// TwinCAT 3 PLC project Tc_SML_MOTION_LAYER
// ProgramVersion: 3.1.4026.18
// libraries:
//   Tc2_Standard, * (Beckhoff Automation GmbH)
//   Tc2_System, * (Beckhoff Automation GmbH)
// project tree:
//   / PlcTask.TcTTO
//   POUs/ MAIN.TcPOU, FB_AxisCtrl.TcPOU, FB_IoLink_In.TcPOU, FB_IoLink_Out.TcPOU, FB_Mapping_In.TcPOU, FB_Mapping_Out.TcPOU, FB_S7RTT_OTG.TcPOU, I_Axis.TcIO, SML_Diagnostics.TcPOU, SML_Home.TcPOU, SML_Power.TcPOU, SML_ProfilePosition.TcPOU, SML_ProfileVelocity.TcPOU, SML_ProfileVelocity_Jog.TcPOU, SML_Reset.TcPOU, SML_Status.TcPOU, SML_Stop.TcPOU, SML_TouchProbe.TcPOU, f_GetProgress.TcPOU, f_GetState.TcPOU
//   DUTs/ E_AXIS_CTRL.TcDUT, E_AXIS_STATE.TcDUT, E_PROGRESS.TcDUT, OpenSML_Axis.TcDUT, SML_DiagCode.TcDUT, ST_AXIS_CTRL.TcDUT, ST_AXIS_INFO.TcDUT, ST_AXIS_STATE.TcDUT, ST_CiA402_Status.TcDUT, ST_DriveIn.TcDUT, ST_DriveOut.TcDUT, ST_MOVE_DATA.TcDUT, U_AXIS_CTRL.TcDUT, U_AXIS_INFO.TcDUT, U_AXIS_STATE.TcDUT, U_MOVE_DATA.TcDUT
//   GVLs/ GVL_SML_CONST.TcGVL

CONFIGURATION Tc_SML_MOTION_LAYER
    RESOURCE PLC ON TwinCAT3
        TASK PlcTask(INTERVAL := T#10ms, PRIORITY := 20);
        PROGRAM MAIN WITH PlcTask : MAIN;
    END_RESOURCE
END_CONFIGURATION

// ---- DUTs/E_AXIS_CTRL.TcDUT
(* ============================================================
   E_AXIS_CTRL - Axis command (eCmd) for FB_AxisCtrl
   SML v6 - Level B (new)

   Level-based command enum: the application writes Ctrl.eCmd;
   FB_AxisCtrl routes the command to the corresponding leaf FB.
   One command at a time => no explicit arbiter (the single value
   of eCmd IS the arbiter).

   Analogous to E_AXIS_CTRL of PLC_MOTION_LAYER, but the commands
   map onto SML's CiA402 FBs instead of the Beckhoff MC_*.
   ============================================================ *)

TYPE E_AXIS_CTRL :
(
    AXIS_NULL          := 0,    // no command: holds the current state
    AXIS_ENABLE        := 1,    // enable drive (Power) and stay idle
    AXIS_DISABLE       := 2,    // disable drive
    AXIS_RESET         := 3,    // fault reset (drive + leaf FBs)
    AXIS_HOME          := 4,    // homing
    AXIS_MOVE_ABS      := 5,    // absolute Profile Position
    AXIS_MOVE_REL      := 6,    // relative Profile Position
    AXIS_MOVE_VELOCITY := 7,    // Profile Velocity (signed velocity)
    AXIS_JOG_POS       := 8,    // jog positive (held)
    AXIS_JOG_NEG       := 9,    // jog negative (held)
    AXIS_MOVE_CSP      := 10,   // CSP (mode 8) + OTG toward Data.lrTargetPosition
    AXIS_STOP          := 11    // Halt (controlled deceleration)
) INT;
END_TYPE

// ---- DUTs/E_AXIS_STATE.TcDUT
(* ============================================================
   E_AXIS_STATE - Axis functional state
   SML v6 - Level B (new)

   Values that are multiples of 100 (= PROGRESS_SPAN) so they can
   compose the COMBINED STATE with E_PROGRESS:
       State.eState = E_AXIS_STATE + E_PROGRESS
   E.g.: AXIS_STATE_MOVING (500) + PROGRESS_BUSY (2) = 502.
   Decompose with f_GetState(502)=500, f_GetProgress(502)=2.

   Here Level B finally USES the f_GetState / f_GetProgress
   functions introduced in Level A.
   ============================================================ *)

TYPE E_AXIS_STATE :
(
    AXIS_STATE_NULL     := 0,     // not initialized
    AXIS_STATE_INIT     := 100,   // init / reset in progress
    AXIS_STATE_DISABLED := 200,   // drive disabled
    AXIS_STATE_IDLE     := 300,   // enabled, stopped, ready
    AXIS_STATE_HOMING   := 400,   // homing
    AXIS_STATE_MOVING   := 500,   // Profile Position / CSP
    AXIS_STATE_VELOCITY := 600,   // Profile Velocity / Jog
    AXIS_STATE_STOPPING := 700,   // Halt
    AXIS_STATE_ERROR    := 900    // error
) INT;
END_TYPE

// ---- DUTs/E_PROGRESS.TcDUT
(* ============================================================
   E_PROGRESS - Unified progress for all SML FBs
   SML v5 - Level A (new)

   Common progress vocabulary, readable by application / HMI /
   diagnostics, replacing the ad-hoc iState:INT semantics used by
   the individual FBs.

   PROJECTION (Level A):
     Each FB keeps its own iState state machine unchanged and, at
     the end of the cycle, exposes eProgress:E_PROGRESS by deriving
     it from iState and from its own flags (xError / xDone / ...).
     No state machine is rewritten.

   COMBINED STATE (Level B groundwork):
     A machine state can be encoded as
       functional_state + E_PROGRESS
     with functional_state a multiple of 100 (see f_GetState /
     f_GetProgress). Not used yet in Level A.
   ============================================================ *)

TYPE E_PROGRESS :
(
    PROGRESS_INVALID := 0,   // not initialized / idle, no request
    PROGRESS_INIT    := 1,   // start request received
    PROGRESS_BUSY    := 2,   // processing
    PROGRESS_PREPARE := 3,   // preparing parameters / preconditions
    PROGRESS_STARTUP := 4,   // running the startup phase
    PROGRESS_CHECK   := 5,   // verifying result / advancing index
    PROGRESS_DONE    := 6,   // completed successfully
    PROGRESS_ERROR   := 7    // error (terminal until reset)
) INT;
END_TYPE

// ---- DUTs/OpenSML_Axis.TcDUT
(* ============================================================
   OpenSML_Axis - Extended CiA402 PDO Data Structure
   SML v4 - Merged from OpenSML + Confa variants

   SOFTWARE STRUCT - no AT %Q*/%I* mapping.
   Use SML_TC3Link to bridge this struct to the TwinCAT I/O tree.
   This keeps the library portable across runtimes and testable
   in simulation without hardware.

   COMPLETE PDO SET (all standard CiA402 objects + Touch Probe):

   OUTPUTS (PLC -> Drive):
     0x6040  ControlWord
     0x6060  Modes_of_operation
     0x607A  Target_Position          [encoder counts]
     0x6081  Profile_Velocity         [drive velocity units - PP mode]
     0x60FF  Target_Velocity          [drive velocity units - PV/CSV mode]
     0x6071  Target_Torque            [0.1 % of rated]
     0x6083  Profile_Acceleration     [drive accel units - PP/PV mode]
     0x6084  Profile_Deceleration     [drive accel units - PP/PV mode]
     0x607C  Home_Offset              [encoder counts - set before homing]
     0x60B8  TouchProbe_ControlWord   [latch trigger control]

   INPUTS (Drive -> PLC):
     0x6041  StatusWord
     0x6061  Modes_of_operation_display
     0x6077  Torque_Actual_Value      [0.1 % of rated]
     0x6064  Position_Actual_Value    [encoder counts]
     0x606C  Velocity_Actual_Value    [drive velocity units]
     0x6078  Current_Actual_Value     [0.1 % of rated]
     0x60F4  Following_Error_Actual_Value [encoder counts]
     0x603F  Error_Code               [drive-specific error number]
     0x60FD  Digital_Inputs           [bitmask of physical digital inputs]
     0x60B9  TouchProbe_StatusWord
     0x60BA  TouchProbe_Rising_Value  [encoder counts - latched on rising edge]
     0x60BB  TouchProbe_Falling_Value [encoder counts - latched on falling edge]

   ControlWord key bits (CiA402 sect. 8.1.3):
     Bit 0  Switch On
     Bit 1  Enable Voltage
     Bit 2  Quick Stop     (1 = run, 0 = activate quick-stop - ACTIVE LOW)
     Bit 3  Enable Operation
     Bit 4  Mode-specific  (New Setpoint in PP / Start Homing in HM)
     Bit 5  Change Setpoint Immediately - blend moves (PP)
     Bit 6  Relative mode  (PP: 0 = absolute, 1 = relative)
     Bit 7  Fault Reset    (rising edge 0->1 clears fault)
     Bit 8  Halt           (1 = decelerate and hold, stay in OperationEnabled)

   StatusWord key bits (CiA402 sect. 8.1.3):
     Bit 0   Ready to Switch On
     Bit 1   Switched On
     Bit 2   Operation Enabled
     Bit 3   Fault
     Bit 4   Voltage Enabled
     Bit 5   Quick Stop     (0 = quick-stop active)
     Bit 6   Switch On Disabled
     Bit 7   Warning
     Bit 9   Remote
     Bit 10  Target Reached / At Velocity / Setpoint Ack (mode-dependent)
     Bit 11  Internal Limit Active
     Bit 12  Mode-specific  (Setpoint Acknowledge in PP / Home Attained in HM)
     Bit 13  Following Error
     Bit 14  Drive-specific (Standstill on many drives)
   ============================================================ *)

TYPE OpenSML_Axis :
STRUCT
    // --- Outputs: PLC -> Drive --------------------------------
    ControlWord          : UINT;   // 0x6040
    Modes_of_operation   : SINT;   // 0x6060
    Target_Position      : DINT;   // 0x607A [encoder counts]
    Profile_Velocity     : UDINT;  // 0x6081 [drive velocity units - PP move speed]
    Target_Velocity      : DINT;   // 0x60FF [drive velocity units - PV/CSV]
    Target_Torque        : INT;    // 0x6071 [0.1 % of rated]
    Profile_Acceleration : UDINT;  // 0x6083 [drive accel units]
    Profile_Deceleration : UDINT;  // 0x6084 [drive accel units]
    Home_Offset          : DINT;   // 0x607C [encoder counts - offset after homing]
    TouchProbe_ControlWord : UINT; // 0x60B8

    // --- Inputs: Drive -> PLC ---------------------------------
    StatusWord                   : UINT;  // 0x6041
    Modes_of_operation_display   : SINT;  // 0x6061
    Torque_Actual_Value          : INT;   // 0x6077 [0.1 % of rated]
    Position_Actual_Value        : DINT;  // 0x6064 [encoder counts]
    Velocity_Actual_Value        : DINT;  // 0x606C [drive velocity units]
    Current_Actual_Value         : INT;   // 0x6078 [0.1 % of rated]
    Following_Error_Actual_Value : DINT;  // 0x60F4 [encoder counts]
    Error_Code                   : UINT;  // 0x603F [drive error number, 0 = no error]
    Digital_Inputs               : UDINT; // 0x60FD [bitmask of physical DI]
    TouchProbe_StatusWord        : UINT;  // 0x60B9
    TouchProbe_Rising_Value      : DINT;  // 0x60BA [encoder counts]
    TouchProbe_Falling_Value     : DINT;  // 0x60BB [encoder counts]
END_STRUCT
END_TYPE

// ---- DUTs/SML_DiagCode.TcDUT
(* ============================================================
   SML_DiagCode - Diagnostic Code Enumeration
   SML v4 - New in v4 (runtime diagnostics)

   Single categorized code used by SML_Diagnostics for both the
   current condition (DiagCode) and the latched first cause
   (FirstFaultCode).  Backed by UINT so it maps cleanly to an HMI
   tag and to alarm tables.

   RANGES:
     0       OK
     1..9    Warnings (motion continues, attention advised)
     10..19  Drive-level faults (CiA402 StatusWord / Error_Code)
     20..29  Library/motion-FB faults (a sub-FB latched an error)
   ============================================================ *)

TYPE SML_DiagCode :
(
    DIAG_OK               := 0,    // No fault, no warning

    // -- Warnings (1..9) ---------------------------------------
    DIAG_WARNING          := 1,    // CiA402 StatusWord bit 7 (generic warning)
    DIAG_INTERNAL_LIMIT   := 2,    // StatusWord bit 11 (internal limit active)

    // -- Drive-level faults (10..19) ---------------------------
    DIAG_DRIVE_FAULT      := 10,   // StatusWord bit 3 (Fault), no specific code
    DIAG_DRIVE_ERRORCODE  := 11,   // StatusWord bit 3 + Error_Code (0x603F) > 0
    DIAG_QUICK_STOP       := 12,   // QuickStopActive (StatusWord bit 5 = 0)
    DIAG_FOLLOWING_ERROR  := 13,   // StatusWord bit 13 (following error)

    // -- Library / motion-FB faults (20..29) -------------------
    DIAG_POWER_ERROR      := 20,   // SML_Power sequence error
    DIAG_HOME_ERROR       := 21,   // SML_Home error (stall/timeout/abort)
    DIAG_MOVE_ERROR       := 22,   // SML_ProfilePosition error (MoveAbs/MoveHome)
    DIAG_VEL_ERROR        := 23,   // SML_ProfileVelocity error
    DIAG_JOG_ERROR        := 24,   // SML_ProfileVelocity_Jog error
    DIAG_TOUCHPROBE_ERROR := 25,   // SML_TouchProbe error
    DIAG_OTG_ERROR        := 26    // FB_S7RTT_OTG constraint error (invalid limits / cycle time)
) UINT;
END_TYPE

// ---- DUTs/ST_AXIS_CTRL.TcDUT
(* ============================================================
   ST_AXIS_CTRL - Command structure (app -> layer)
   SML v6 - Level B (new)

   The "Ctrl" data contract of the Motion Layer pattern. A flat,
   serializable structure (no pointer/interface inside): accessible
   via ADS symbol or copyable onto a bus (MAPPING groundwork).

   The eCmd command is level-based. Motion parameters live in
   ST_MOVE_DATA ("Data").
   ============================================================ *)

TYPE ST_AXIS_CTRL :
STRUCT
    eCmd           : E_AXIS_CTRL;        // requested command
    xEmergencyStop : BOOL := TRUE;       // TRUE = run / FALSE = quick-stop (CiA402 bit 2)
    xSimulation    : BOOL;               // mirror Target_Position -> Position_Actual_Value

    // -- configuration (rarely changed) -----------------------
    Scale          : LREAL := 4096.0;    // [counts/unit] - must be > 0
    CycleTime      : LREAL := 0.001;     // [s] - must match the task (OTG)
    PositionWindow : LREAL := 0.01;      // in-position deadband [units]
    HomeOffset     : DINT  := 0;         // homing offset [encoder counts] -> 0x607C

    // -- TouchProbe (parallel to motion, not an eCmd) ----------
    xTouchProbeEnable  : BOOL;           // arm the TouchProbe hardware
    xTouchProbeRising  : BOOL;           // arm the latch on the rising edge
    xTouchProbeFalling : BOOL;           // arm the latch on the falling edge
END_STRUCT
END_TYPE

// ---- DUTs/ST_AXIS_INFO.TcDUT
(* ============================================================
   ST_AXIS_INFO - Info structure (layer -> app)
   SML v6 - Level B (new)

   The "Info" data contract. Actual values and axis status bits,
   in user units.
   ============================================================ *)

TYPE ST_AXIS_INFO :
STRUCT
    lrActualPosition : LREAL;    // actual position [units]
    lrActualVelocity : LREAL;    // actual velocity [units/s]
    xEnabled         : BOOL;     // drive in OperationEnabled
    xHomed           : BOOL;     // homing done at least once (latch)
    xMoving          : BOOL;     // axis is moving
    xInPosition      : BOOL;     // within PositionWindow (CSP path)

    // -- full CiA402 decoder (from SML_Status) -----------------
    Status           : ST_CiA402_Status;

    // -- TouchProbe results (from SML_TouchProbe) --------------
    xTouchProbeDoneR       : BOOL;
    xTouchProbeDoneF       : BOOL;
    xTouchProbeBusy        : BOOL;
    xTouchProbeError       : BOOL;
    TouchProbeRisingValue  : DINT;   // [encoder counts]
    TouchProbeFallingValue : DINT;   // [encoder counts]
END_STRUCT
END_TYPE

// ---- DUTs/ST_AXIS_STATE.TcDUT
(* ============================================================
   ST_AXIS_STATE - State structure (layer -> app)
   SML v6 - Level B (new)

   The "State" data contract. Command result + progress.
   eState is the COMBINED STATE (E_AXIS_STATE + E_PROGRESS);
   use f_GetState / f_GetProgress to decompose it.
   ============================================================ *)

TYPE ST_AXIS_STATE :
STRUCT
    eState         : INT;            // combined state = E_AXIS_STATE + E_PROGRESS
    eProgress      : E_PROGRESS;     // progress (handy, already decomposed)
    eCmdActive     : E_AXIS_CTRL;    // command being executed
    xDone          : BOOL;           // current command complete
    xError         : BOOL;           // aggregated error

    // -- diagnostics (from SML_Diagnostics) -------------------
    DiagCode       : SML_DiagCode;
    DiagText       : STRING(80);
    FirstFaultCode : SML_DiagCode;
    FirstFaultText : STRING(80);
END_STRUCT
END_TYPE

// ---- DUTs/ST_CiA402_Status.TcDUT
(* ============================================================
   ST_CiA402_Status - Full CiA402 status decoder
   SML v9 - Level B (new)

   Mirrors the outputs of the SML_Status decoder, made available in
   the data contract as a sub-struct of ST_AXIS_INFO (Info.Status).
   Brings into FB_AxisCtrl the granular status bits that used to be
   exposed only by FB_SML.
   ============================================================ *)

TYPE ST_CiA402_Status :
STRUCT
    // -- CiA402 state machine ----------------------------------
    NotReadyToSwitchOn  : BOOL;
    SwitchOnDisabled    : BOOL;
    ReadyToSwitchOn     : BOOL;
    SwitchedOn          : BOOL;
    OperationEnabled    : BOOL;
    QuickStopActive     : BOOL;
    FaultReactionActive : BOOL;
    Fault               : BOOL;

    // -- general status ----------------------------------------
    Warning             : BOOL;   // bit 7
    TargetReached       : BOOL;   // bit 10 (mode-dependent)
    Halted              : BOOL;
    VoltageEnabled      : BOOL;   // bit 4
    InternalLimit       : BOOL;   // bit 11

    // -- active operating mode ---------------------------------
    ProfilePositionMode : BOOL;   // 1
    ProfileVelocityMode : BOOL;   // 3
    VelocityMode        : BOOL;   // 2 (legacy)
    TorqueProfileMode   : BOOL;   // 4
    HomingMode          : BOOL;   // 6
    SyncPositionMode    : BOOL;   // 8 (CSP)
    SyncVelocityMode    : BOOL;   // 9 (CSV)

    // -- motion ------------------------------------------------
    Moving              : BOOL;
    StandStill          : BOOL;
    Homed               : BOOL;

    // -- error / detail ----------------------------------------
    Err                 : BOOL;   // Error_Code != 0
    ErrId               : UINT;   // 0x603F
    ActTorque           : INT;    // 0x6077 [0.1% of rated]
    FollowingError      : DINT;   // 0x60F4 [encoder counts]
END_STRUCT
END_TYPE

// ---- DUTs/ST_DriveIn.TcDUT
(* ============================================================
   ST_DriveIn - INPUT process image (Drive -> PLC)
   SML v9 - I/O bridge (new)

   The "input" half of OpenSML_Axis, SAME order and same types.
   Used for the I/O bridge: declared AT %I* (mapped to the drive's
   TxPDOs) and copied into GVL_AXIS.Axis[n] before the computation.

   Valid for both CoDeSys and TwinCAT (generic IEC 61131-3 ST).
   ============================================================ *)

TYPE ST_DriveIn :
STRUCT
    StatusWord                   : UINT;   // 0x6041
    Modes_of_operation_display   : SINT;   // 0x6061
    Torque_Actual_Value          : INT;    // 0x6077 [0.1 % rated]
    Position_Actual_Value        : DINT;   // 0x6064 [encoder counts]
    Velocity_Actual_Value        : DINT;   // 0x606C [drive velocity units]
    Current_Actual_Value         : INT;    // 0x6078 [0.1 % rated]
    Following_Error_Actual_Value : DINT;   // 0x60F4 [encoder counts]
    Error_Code                   : UINT;   // 0x603F [0 = no error]
    Digital_Inputs               : UDINT;  // 0x60FD [DI bitmask]
    TouchProbe_StatusWord        : UINT;   // 0x60B9
    TouchProbe_Rising_Value      : DINT;   // 0x60BA [encoder counts]
    TouchProbe_Falling_Value     : DINT;   // 0x60BB [encoder counts]
END_STRUCT
END_TYPE

// ---- DUTs/ST_DriveOut.TcDUT
(* ============================================================
   ST_DriveOut - OUTPUT process image (PLC -> Drive)
   SML v9 - I/O bridge (new)

   The "output" half of OpenSML_Axis, SAME order and same types.
   Used for the I/O bridge: declared AT %Q* (mapped to the drive's
   RxPDOs) and copied from GVL_AXIS.Axis[n] after the computation.

   Valid for both CoDeSys and TwinCAT (generic IEC 61131-3 ST).
   On CoDeSys, as an alternative, you can directly link
   GVL_AXIS.Axis[n].<member> in the I/O Mapping tab (no bridge).
   ============================================================ *)

TYPE ST_DriveOut :
STRUCT
    ControlWord            : UINT;   // 0x6040
    Modes_of_operation     : SINT;   // 0x6060
    Target_Position        : DINT;   // 0x607A [encoder counts]
    Profile_Velocity       : UDINT;  // 0x6081 [drive velocity units - PP]
    Target_Velocity        : DINT;   // 0x60FF [drive velocity units - PV/CSV]
    Target_Torque          : INT;    // 0x6071 [0.1 % rated]
    Profile_Acceleration   : UDINT;  // 0x6083 [drive accel units]
    Profile_Deceleration   : UDINT;  // 0x6084 [drive accel units]
    Home_Offset            : DINT;   // 0x607C [encoder counts]
    TouchProbe_ControlWord : UINT;   // 0x60B8
END_STRUCT
END_TYPE

// ---- DUTs/ST_MOVE_DATA.TcDUT
(* ============================================================
   ST_MOVE_DATA - Setpoints and dynamic limits (app -> layer)
   SML v6 - Level B (new)

   The "Data" data contract. All values are in USER UNITS (LREAL).
   FB_AxisCtrl converts to the drive's raw units via Ctrl.Scale
   before passing them to the leaf FBs (PP/PV/Jog); the CSP/OTG
   path works directly in user units.

   Scaling note: velocity/acceleration scale is assumed equal to
   position scale (multiply by Scale). For drives whose velocity
   units 0x6081/0x60FF differ, refine the conversion in the FB.
   ============================================================ *)

TYPE ST_MOVE_DATA :
STRUCT
    lrTargetPosition : LREAL;              // target [units] for MOVE_ABS/REL/CSP
    lrVelocity       : LREAL := 10.0;      // velocity [units/s]; signed for MOVE_VELOCITY
    lrAcceleration   : LREAL := 1000.0;    // [units/s^2]
    lrDeceleration   : LREAL := 1000.0;    // [units/s^2]
    lrJerk           : LREAL := 10000.0;   // [units/s^3] - CSP/OTG only
END_STRUCT
END_TYPE

// ---- DUTs/U_AXIS_CTRL.TcDUT
(* ============================================================
   U_AXIS_CTRL - Bus UNION for the axis command
   SML v8 - Level B / MAPPING (new)

   Overlay of the same memory block as:
     - stData : ST_AXIS_CTRL   (typed view for the logic)
     - aRaw   : byte block      (raw view for fieldbus mapping)

   Fixed size = MAP_SIZE_CTRL (>= SIZEOF(ST_AXIS_CTRL), checked by
   FB_Mapping_In). Lets you link the element to the process image as
   a struct or as a raw block without changing the mapped size.
   ============================================================ *)

TYPE U_AXIS_CTRL :
UNION
    stData : ST_AXIS_CTRL;
    aRaw   : ARRAY[1..GVL_SML_CONST.MAP_SIZE_CTRL] OF BYTE;
END_UNION
END_TYPE

// ---- DUTs/U_AXIS_INFO.TcDUT
(* ============================================================
   U_AXIS_INFO - Bus UNION for the axis info
   SML v8 - Level B / MAPPING (new)

   stData : ST_AXIS_INFO (typed) / aRaw : byte block (fieldbus).
   Fixed size = MAP_SIZE_INFO (>= SIZEOF(ST_AXIS_INFO)).
   ============================================================ *)

TYPE U_AXIS_INFO :
UNION
    stData : ST_AXIS_INFO;
    aRaw   : ARRAY[1..GVL_SML_CONST.MAP_SIZE_INFO] OF BYTE;
END_UNION
END_TYPE

// ---- DUTs/U_AXIS_STATE.TcDUT
(* ============================================================
   U_AXIS_STATE - Bus UNION for the axis state
   SML v8 - Level B / MAPPING (new)

   stData : ST_AXIS_STATE (typed) / aRaw : byte block (fieldbus).
   Fixed size = MAP_SIZE_STATE (>= SIZEOF(ST_AXIS_STATE)).
   ============================================================ *)

TYPE U_AXIS_STATE :
UNION
    stData : ST_AXIS_STATE;
    aRaw   : ARRAY[1..GVL_SML_CONST.MAP_SIZE_STATE] OF BYTE;
END_UNION
END_TYPE

// ---- DUTs/U_MOVE_DATA.TcDUT
(* ============================================================
   U_MOVE_DATA - Bus UNION for the motion setpoints
   SML v8 - Level B / MAPPING (new)

   stData : ST_MOVE_DATA (typed) / aRaw : byte block (fieldbus).
   Fixed size = MAP_SIZE_DATA (>= SIZEOF(ST_MOVE_DATA)).
   ============================================================ *)

TYPE U_MOVE_DATA :
UNION
    stData : ST_MOVE_DATA;
    aRaw   : ARRAY[1..GVL_SML_CONST.MAP_SIZE_DATA] OF BYTE;
END_UNION
END_TYPE

// ---- GVLs/GVL_SML_CONST.TcGVL
(* ============================================================
   GVL_SML_CONST - LIBRARY constants (invariants)
   SML

   Only constants owned by the library (machine-independent).
   The application configuration (number of axes) lives in GVL_App.MAX_AXIS.
   Qualified reference: GVL_SML_CONST.PROGRESS_SPAN, ...
   ============================================================ *)

{attribute 'qualified_only'}
VAR_GLOBAL CONSTANT
    PROGRESS_SPAN : DINT := 100;   // progress band width in the combined state
                                   // (E_AXIS_STATE values are multiples of this)

    // -- MAPPING: fixed size (bytes) of the bus blocks for the UNIONs --
    // Must be >= SIZEOF of the corresponding struct (checked at runtime
    // by FB_Mapping_In/Out via Check). Fixed for a stable process image
    // on the fieldbus.
    MAP_SIZE_CTRL  : UDINT := 64;    // >= SIZEOF(ST_AXIS_CTRL)
    MAP_SIZE_DATA  : UDINT := 64;    // >= SIZEOF(ST_MOVE_DATA)
    MAP_SIZE_STATE : UDINT := 256;   // >= SIZEOF(ST_AXIS_STATE) (holds 2x STRING(80))
    MAP_SIZE_INFO  : UDINT := 128;   // >= SIZEOF(ST_AXIS_INFO) (with Status + TouchProbe)
END_VAR

// ---- POUs/I_Axis.TcIO
INTERFACE I_Axis

METHOD Enable : E_PROGRESS
VAR_INPUT
END_VAR
END_METHOD

METHOD Disable : E_PROGRESS
VAR_INPUT
END_VAR
END_METHOD

METHOD Reset : E_PROGRESS
VAR_INPUT
END_VAR
END_METHOD

METHOD Home : E_PROGRESS
VAR_INPUT
END_VAR
END_METHOD

METHOD MoveAbsolute : E_PROGRESS
VAR_INPUT
    lrPosition : LREAL;   // [units]
    lrVelocity : LREAL;   // [units/s]
END_VAR
END_METHOD

METHOD MoveRelative : E_PROGRESS
VAR_INPUT
    lrDistance : LREAL;   // [units]
    lrVelocity : LREAL;   // [units/s]
END_VAR
END_METHOD

METHOD MoveVelocity : E_PROGRESS
VAR_INPUT
    lrVelocity : LREAL;   // [units/s] signed
END_VAR
END_METHOD

METHOD Jog : E_PROGRESS
VAR_INPUT
    xForward   : BOOL;
    xReverse   : BOOL;
    lrVelocity : LREAL;   // magnitude [units/s]
END_VAR
END_METHOD

METHOD MoveFollow : E_PROGRESS
VAR_INPUT
    lrPosition : LREAL;   // [units] - online re-targetable
    lrVelocity : LREAL;   // [units/s]
END_VAR
END_METHOD

METHOD Stop : E_PROGRESS
VAR_INPUT
END_VAR
END_METHOD

PROPERTY Position : LREAL
GET
END_GET
END_PROPERTY

PROPERTY Enabled : BOOL
GET
END_GET
END_PROPERTY

END_INTERFACE

// ---- POUs/MAIN.TcPOU
PROGRAM MAIN
VAR
END_VAR

END_PROGRAM

// ---- POUs/FB_Mapping_In.TcPOU
(* ============================================================
   FB_Mapping_In - MAPPING bridge FB: bus -> internal (command)
   SML - Level B / MAPPING (library FB)

   Copies the command/setpoint from the bus UNIONs into the internal
   Ctrl/Data structs, for all axes:
     CtrlBus[].stData -> Ctrl[]   ,   DataBus[].stData -> Data[]
   Call at the START of the task, before the axis loop.

   Reusable: arrays passed by VAR_IN_OUT as ARRAY[*] (variable
   length) - no dependency on MAX_AXIS or on any application GVL. The
   application keeps the bus UNION arrays (e.g. GVL_AXIS_MAP.Ctrl/Data)
   and its enable flag, and instantiates this FB.

   GATE: copies only when xEnable = TRUE.
   Runtime size check: if a struct exceeds its bus block (MAP_SIZE_CTRL/DATA),
   the copy is blocked for safety (resize MAP_SIZE_* in GVL_SML_CONST).
   Precondition: all arrays have the same bounds (one entry per axis).
   ============================================================ *)

FUNCTION_BLOCK FB_Mapping_In
VAR_INPUT
    xEnable : BOOL;   // TRUE = perform the copy; FALSE = bypass
END_VAR
VAR_IN_OUT
    CtrlBus : ARRAY[*] OF U_AXIS_CTRL;   // <- bus command  (.stData)
    DataBus : ARRAY[*] OF U_MOVE_DATA;   // <- bus setpoint (.stData)
    Ctrl    : ARRAY[*] OF ST_AXIS_CTRL;  // -> internal command
    Data    : ARRAY[*] OF ST_MOVE_DATA;  // -> internal setpoint
END_VAR
VAR
    i       : DINT;
    bSizeOk : BOOL;
END_VAR

IF NOT xEnable THEN RETURN; END_IF

// -- Bus block size check (safety) ----------------------------
bSizeOk := (SIZEOF(ST_AXIS_CTRL) <= GVL_SML_CONST.MAP_SIZE_CTRL)
       AND (SIZEOF(ST_MOVE_DATA) <= GVL_SML_CONST.MAP_SIZE_DATA);
IF NOT bSizeOk THEN RETURN; END_IF   // blocked: resize MAP_SIZE_*

// -- Copy bus -> internal -------------------------------------
FOR i := LOWER_BOUND(Ctrl, 1) TO UPPER_BOUND(Ctrl, 1) DO
    Ctrl[i] := CtrlBus[i].stData;
    Data[i] := DataBus[i].stData;
END_FOR

END_FUNCTION_BLOCK

// ---- POUs/FB_AxisCtrl.TcPOU
(* ============================================================
   FB_AxisCtrl - Command-driven axis control FB (Level B)
   SML v6 - new

   Brings the Motion Layer pattern of PLC_MOTION_LAYER onto SML:
   instead of wrapping the Beckhoff MC_*, this FB drives DIRECTLY
   SML's CiA402 leaf FBs (Power/Home/ProfilePosition/ProfileVelocity/
   Jog/Stop) + the CSP path with FB_S7RTT_OTG.

   SUPERSET of FB_SML (v9): it also integrates the full status decoder
   SML_Status (-> Info.Status, all CiA402 bits) and SML_TouchProbe
   (-> Info.xTouchProbe* fields, commanded via Ctrl.xTouchProbe* inputs). The TouchProbe
   is PARALLEL to motion (it is not an eCmd) and its error feeds the
   diagnostics but NOT the combined motion state (eState).

   INPUTS / OUTPUTS via the data contract (VAR_IN_OUT):
     Axis  : OpenSML_Axis   drive PDO image
     Ctrl  : ST_AXIS_CTRL   command (eCmd) + config             (app -> layer)
     Data  : ST_MOVE_DATA   motion setpoints [user units]       (app -> layer)
     State : ST_AXIS_STATE  result + combined state            (layer -> app)
     Info  : ST_AXIS_INFO   actual values + bits                (layer -> app)

   ARBITRATION: eCmd is a single value => only one motion command
   active per cycle. No explicit arbiter (unlike FB_SML).

   ENTRY-POINT: call cyclically. As an alternative to writing
   Ctrl.eCmd, you can use the I_Axis methods (equivalent setters).

   IMPLEMENTS I_Axis.
   ============================================================ *)

FUNCTION_BLOCK FB_AxisCtrl IMPLEMENTS I_Axis
VAR_IN_OUT
    Axis  : OpenSML_Axis;
    Ctrl  : ST_AXIS_CTRL;
    Data  : ST_MOVE_DATA;
    State : ST_AXIS_STATE;
    Info  : ST_AXIS_INFO;
END_VAR
VAR
    // -- leaf FBs (execution level, in place of the MC_*) ------
    inst_Power   : SML_Power;
    inst_Reset   : SML_Reset;
    inst_Home    : SML_Home;
    inst_MoveAbs : SML_ProfilePosition;
    inst_MoveVel : SML_ProfileVelocity;
    inst_Jog     : SML_ProfileVelocity_Jog;
    inst_Stop       : SML_Stop;
    inst_Diag       : SML_Diagnostics;
    inst_Status     : SML_Status;         // full CiA402 decoder (superset of FB_SML)
    inst_TouchProbe : SML_TouchProbe;     // TouchProbe (parallel to motion)
    otg          : FB_S7RTT_OTG;

    // -- command -----------------------------------------------
    _eCmd, _eCmdOld : E_AXIS_CTRL;

    // -- latch / pulse ----------------------------------------
    _bEnableReq  : BOOL;       // enable request (ENABLE/DISABLE)
    _xReset      : BOOL;       // reset active (level)
    _xHomedLatch : BOOL;       // homing done at least once
    _eCspState   : INT;        // CSP sub-state: 0 seed, 1 run

    // -- unit conversions (user -> raw drive) -----------------
    _diPos   : DINT;
    _diVelSg : DINT;           // signed velocity (PV)
    _diVelMg : DINT;           // magnitude (Jog)
    _udiVel  : UDINT;
    _udiAcc  : UDINT;
    _udiDec  : UDINT;

    // -- gate -------------------------------------------------
    _xMotionEnable : BOOL;

    // -- flags from the leaf FBs ------------------------------
    _xEnabled, _xPowerErr                          : BOOL;
    _xResetDone, _xResetErr                        : BOOL;
    _xHomeBusy, _xHomeDone, _xHomeErr              : BOOL;
    _xMoveDone, _xMoveBusy, _xMoveMoving, _xMoveErr: BOOL;
    _xAtVel, _xVelMoving, _xVelErr                 : BOOL;
    _xJogMoving, _xJogErr                          : BOOL;
    _xStopped                                      : BOOL;
    _xTpErr                                        : BOOL;   // TouchProbe error (parallel)
    _xInPos, _xCspErr                              : BOOL;
    _xActiveFault, _xAnyErr                        : BOOL;

    // -- combined-state computation ---------------------------
    _eBase : E_AXIS_STATE;
    _eProg : E_PROGRESS;
END_VAR

//------------------------------------------------------------------------------
// /input + guards
//------------------------------------------------------------------------------
_eCmd := Ctrl.eCmd;

IF Ctrl.Scale = 0.0 THEN Ctrl.Scale := 1.0; END_IF   // divide-by-zero guard

IF Ctrl.xSimulation THEN
    Axis.Position_Actual_Value := Axis.Target_Position;  // mirror in simulation
END_IF

// enable latch: any command != NULL/DISABLE implies enable
IF    _eCmd = AXIS_DISABLE THEN _bEnableReq := FALSE;
ELSIF _eCmd <> AXIS_NULL   THEN _bEnableReq := TRUE;
END_IF

_xReset        := (_eCmd = AXIS_RESET);
_xMotionEnable := _xEnabled AND Ctrl.xEmergencyStop;

// user units -> drive raw units (see scaling note in ST_MOVE_DATA)
_diPos   := LREAL_TO_DINT (Data.lrTargetPosition * Ctrl.Scale);
_diVelSg := LREAL_TO_DINT (Data.lrVelocity       * Ctrl.Scale);
_diVelMg := LREAL_TO_DINT (ABS(Data.lrVelocity)  * Ctrl.Scale);
_udiVel  := LREAL_TO_UDINT(ABS(Data.lrVelocity)  * Ctrl.Scale);
_udiAcc  := LREAL_TO_UDINT(Data.lrAcceleration   * Ctrl.Scale);
_udiDec  := LREAL_TO_UDINT(Data.lrDeceleration   * Ctrl.Scale);
//------------------------------------------------------------------------------
// input + guards/
//------------------------------------------------------------------------------

//------------------------------------------------------------------------------
// /leaf FBs - called every cycle, gated via eCmd (like FB_SML)
//------------------------------------------------------------------------------
inst_Power(
    Axis           := Axis,
    xExecute       := _bEnableReq,
    xEmergencyStop := Ctrl.xEmergencyStop,
    xDone          => _xEnabled,
    xError         => _xPowerErr);

inst_Reset(
    Axis     := Axis,
    xExecute := _xReset,
    xDone    => _xResetDone,
    xError   => _xResetErr);

inst_Home(
    Axis         := Axis,
    xEnable      := _xMotionEnable,
    xExecute     := (_eCmd = AXIS_HOME),
    xReset       := _xReset,
    diHomeOffset := Ctrl.HomeOffset,
    xBusy        => _xHomeBusy,
    xDone        => _xHomeDone,
    xError       => _xHomeErr);
IF _xHomeDone THEN _xHomedLatch := TRUE; END_IF

inst_MoveAbs(
    Axis                   := Axis,
    xEnable                := _xMotionEnable,
    xExecute               := (_eCmd = AXIS_MOVE_ABS) OR (_eCmd = AXIS_MOVE_REL),
    xReset                 := _xReset,
    xContinueMove          := FALSE,
    xRelativeMode          := (_eCmd = AXIS_MOVE_REL),
    diTargetPosition       := _diPos,
    udiProfileVelocity     := _udiVel,
    udiProfileAcceleration := _udiAcc,
    udiProfileDeceleration := _udiDec,
    xDone                  => _xMoveDone,
    xBusy                  => _xMoveBusy,
    xMoving                => _xMoveMoving,
    xError                 => _xMoveErr);

inst_MoveVel(
    Axis                   := Axis,
    xEnable                := _xMotionEnable,
    xExecute               := (_eCmd = AXIS_MOVE_VELOCITY),
    xReset                 := _xReset,
    diTargetVelocity       := _diVelSg,
    udiProfileAcceleration := _udiAcc,
    udiProfileDeceleration := _udiDec,
    xMoving                => _xVelMoving,
    xAtVelocity            => _xAtVel,
    xError                 => _xVelErr);

inst_Jog(
    Axis                   := Axis,
    xEnable                := _xMotionEnable,
    xExecute_Jog_F         := (_eCmd = AXIS_JOG_POS),
    xExecute_Jog_R         := (_eCmd = AXIS_JOG_NEG),
    xReset                 := _xReset,
    diProfileVelocity      := _diVelMg,
    udiProfileAcceleration := _udiAcc,
    udiProfileDeceleration := _udiDec,
    xMoving                => _xJogMoving,
    xError                 => _xJogErr);

inst_Stop(
    Axis     := Axis,
    xStop    := (_eCmd = AXIS_STOP),
    xStopped => _xStopped);

// full CiA402 decoder (read-only) -> Info.Status
inst_Status(
    Axis                       := Axis,
    xEnable                    := TRUE,
    Status_NotReadyToSwitchOn  => Info.Status.NotReadyToSwitchOn,
    Status_SwitchOnDisabled    => Info.Status.SwitchOnDisabled,
    Status_ReadyToSwitchOn     => Info.Status.ReadyToSwitchOn,
    Status_SwitchedOn          => Info.Status.SwitchedOn,
    Status_OperationEnabled    => Info.Status.OperationEnabled,
    Status_QuickStopActive     => Info.Status.QuickStopActive,
    Status_FaultReactionActive => Info.Status.FaultReactionActive,
    Status_Fault               => Info.Status.Fault,
    Status_Warning             => Info.Status.Warning,
    Status_TargetReached       => Info.Status.TargetReached,
    Status_Halted              => Info.Status.Halted,
    Status_VoltageEnabled      => Info.Status.VoltageEnabled,
    Status_InternalLimit       => Info.Status.InternalLimit,
    Status_ProfilePositionMode => Info.Status.ProfilePositionMode,
    Status_ProfileVelocityMode => Info.Status.ProfileVelocityMode,
    Status_VelocityMode        => Info.Status.VelocityMode,
    Status_TorqueProfileMode   => Info.Status.TorqueProfileMode,
    Status_HomingMode          => Info.Status.HomingMode,
    Status_SyncPositionMode    => Info.Status.SyncPositionMode,
    Status_SyncVelocityMode    => Info.Status.SyncVelocityMode,
    Status_Moving              => Info.Status.Moving,
    Status_StandStill          => Info.Status.StandStill,
    Status_Homed               => Info.Status.Homed,
    StatusErr                  => Info.Status.Err,
    ErrId                      => Info.Status.ErrId,
    ActPosition                => ,
    ActSpeed                   => ,
    ActTorque                  => Info.Status.ActTorque,
    FollowingError             => Info.Status.FollowingError);

// TouchProbe (parallel to motion) -> Info.xTouchProbe*
inst_TouchProbe(
    Axis                     := Axis,
    xEnable                  := _xMotionEnable,
    xExecute                 := Ctrl.xTouchProbeEnable,
    xRisingCapture           := Ctrl.xTouchProbeEnable AND Ctrl.xTouchProbeRising,
    xFallingCapture          := Ctrl.xTouchProbeEnable AND Ctrl.xTouchProbeFalling,
    xReset                   := _xReset,
    xDone_R                  => Info.xTouchProbeDoneR,
    xDone_F                  => Info.xTouchProbeDoneF,
    xBusy                    => Info.xTouchProbeBusy,
    xError                   => _xTpErr,
    TouchProbe_Rising_Value  => Info.TouchProbeRisingValue,
    TouchProbe_Falling_Value => Info.TouchProbeFallingValue);
Info.xTouchProbeError := _xTpErr;
//------------------------------------------------------------------------------
// leaf FBs/
//------------------------------------------------------------------------------

//------------------------------------------------------------------------------
// /CSP + OTG - active only with eCmd = AXIS_MOVE_CSP
//------------------------------------------------------------------------------
_xInPos := FALSE;
IF (_eCmd = AXIS_MOVE_CSP) AND _xMotionEnable THEN
    Info.lrActualPosition := DINT_TO_LREAL(Axis.Position_Actual_Value) / Ctrl.Scale;
    CASE _eCspState OF
        0: // switch to CSP (mode 8) + seed OTG at the actual position
            Axis.Modes_of_operation := 8;
            Axis.ControlWord.3      := (Axis.Modes_of_operation_display = 8);
            otg(
                xInit            := TRUE,
                CurrentPosition  := Info.lrActualPosition,
                ControlInterface := TRUE,
                TargetPosition   := Data.lrTargetPosition,
                TargetVelocity   := 0.0,
                CycleTIme        := Ctrl.CycleTime,
                MaxVelocity      := Data.lrVelocity,
                MaxAcceleration  := Data.lrAcceleration,
                MaxJerk          := Data.lrJerk);
            IF (Axis.StatusWord.2 AND Axis.Modes_of_operation_display = 8) OR Ctrl.xSimulation THEN
                _eCspState := 1;
            END_IF

        1: // CSP motion loop
            otg(
                xInit            := FALSE,
                ControlInterface := FALSE,
                TargetPosition   := Data.lrTargetPosition,
                TargetVelocity   := 0.0,
                CycleTIme        := Ctrl.CycleTime,
                MaxVelocity      := Data.lrVelocity,
                MaxAcceleration  := Data.lrAcceleration,
                MaxJerk          := Data.lrJerk);
            Axis.Target_Position := LREAL_TO_DINT(otg.NewPosition * Ctrl.Scale);
            _xInPos := ABS(otg.NewPosition - Data.lrTargetPosition) < Ctrl.PositionWindow;
    END_CASE
    _xCspErr := Axis.StatusWord.13 OR Axis.StatusWord.3 OR otg.xError OR _xPowerErr;
ELSE
    _eCspState := 0;      // reset the sub-state when not in CSP
    _xCspErr   := FALSE;
END_IF
//------------------------------------------------------------------------------
// CSP + OTG/
//------------------------------------------------------------------------------

//------------------------------------------------------------------------------
// /aggregated diagnostics
//------------------------------------------------------------------------------
inst_Diag(
    Axis             := Axis,
    xReset           := _xReset,
    xResetCount      := FALSE,
    xPowerError      := _xPowerErr,
    xHomeError       := _xHomeErr,
    xMoveError       := _xMoveErr,
    xVelError        := _xVelErr,
    xJogError        := _xJogErr,
    xTouchProbeError := _xTpErr,
    xOtgError        := otg.xError,
    DiagCode         => State.DiagCode,
    DiagText         => State.DiagText,
    xActiveFault     => _xActiveFault,
    xActiveWarning   => ,
    FirstFaultCode   => State.FirstFaultCode,
    FirstFaultText   => State.FirstFaultText,
    DriveErrorCode   => ,
    FollowingError   => ,
    FaultCount       => );
//------------------------------------------------------------------------------
// aggregated diagnostics/
//------------------------------------------------------------------------------

//------------------------------------------------------------------------------
// /Info (feedback) + aggregated error
//------------------------------------------------------------------------------
Info.lrActualPosition := DINT_TO_LREAL(Axis.Position_Actual_Value) / Ctrl.Scale;
Info.lrActualVelocity := DINT_TO_LREAL(Axis.Velocity_Actual_Value) / Ctrl.Scale;
Info.xEnabled         := _xEnabled;
Info.xHomed           := _xHomedLatch;
Info.xMoving          := _xMoveMoving OR _xVelMoving OR _xJogMoving OR (_eCmd = AXIS_MOVE_CSP);
Info.xInPosition      := _xInPos;

_xAnyErr := _xPowerErr OR _xHomeErr OR _xMoveErr OR _xVelErr
            OR _xJogErr OR _xCspErr OR _xResetErr;
//------------------------------------------------------------------------------
// Info + error/
//------------------------------------------------------------------------------

//------------------------------------------------------------------------------
// /combined state  eState = E_AXIS_STATE + E_PROGRESS
//------------------------------------------------------------------------------
IF _xAnyErr THEN
    _eBase := AXIS_STATE_ERROR;
    _eProg := PROGRESS_ERROR;
ELSE
    CASE _eCmd OF
        AXIS_NULL:
            IF _xEnabled THEN _eBase := AXIS_STATE_IDLE; ELSE _eBase := AXIS_STATE_DISABLED; END_IF
            _eProg := PROGRESS_INVALID;

        AXIS_ENABLE:
            _eBase := AXIS_STATE_IDLE;
            IF _xEnabled THEN _eProg := PROGRESS_DONE; ELSE _eProg := PROGRESS_BUSY; END_IF

        AXIS_DISABLE:
            _eBase := AXIS_STATE_DISABLED;
            IF _xEnabled THEN _eProg := PROGRESS_BUSY; ELSE _eProg := PROGRESS_DONE; END_IF

        AXIS_RESET:
            _eBase := AXIS_STATE_INIT;
            IF _xResetDone THEN _eProg := PROGRESS_DONE; ELSE _eProg := PROGRESS_BUSY; END_IF

        AXIS_HOME:
            _eBase := AXIS_STATE_HOMING;
            IF _xHomeDone THEN _eProg := PROGRESS_DONE; ELSE _eProg := PROGRESS_BUSY; END_IF

        AXIS_MOVE_ABS, AXIS_MOVE_REL:
            _eBase := AXIS_STATE_MOVING;
            IF _xMoveDone THEN _eProg := PROGRESS_DONE; ELSE _eProg := PROGRESS_BUSY; END_IF

        AXIS_MOVE_CSP:
            _eBase := AXIS_STATE_MOVING;
            IF _xInPos THEN _eProg := PROGRESS_DONE; ELSE _eProg := PROGRESS_BUSY; END_IF

        AXIS_MOVE_VELOCITY:
            _eBase := AXIS_STATE_VELOCITY;
            IF _xAtVel THEN _eProg := PROGRESS_DONE; ELSE _eProg := PROGRESS_BUSY; END_IF

        AXIS_JOG_POS, AXIS_JOG_NEG:
            _eBase := AXIS_STATE_VELOCITY;
            _eProg := PROGRESS_BUSY;      // continuous jog: no discrete DONE

        AXIS_STOP:
            _eBase := AXIS_STATE_STOPPING;
            IF _xStopped THEN _eProg := PROGRESS_DONE; ELSE _eProg := PROGRESS_BUSY; END_IF
    END_CASE
END_IF

State.eProgress  := _eProg;
State.eState     := TO_INT(_eBase) + TO_INT(_eProg);   // combined state
State.eCmdActive := _eCmd;
State.xError     := _xAnyErr;
State.xDone      := (_eProg = PROGRESS_DONE);

_eCmdOld := _eCmd;
//------------------------------------------------------------------------------
// combined state/
//------------------------------------------------------------------------------


(* ============================================================
   METHODS / PROPERTIES of I_Axis
   Real code in  FB_AxisCtrl_METHODS.txt  (to be created as
   METHOD/PROPERTY objects under this FB in CoDeSys).
   They are setters: they set Ctrl.eCmd (+ Data) and return
   State.eProgress.
   ============================================================ *)

METHOD Enable : E_PROGRESS
VAR_INPUT
END_VAR
Ctrl.eCmd := AXIS_ENABLE;
Enable    := State.eProgress;
END_METHOD

METHOD Disable : E_PROGRESS
VAR_INPUT
END_VAR
Ctrl.eCmd := AXIS_DISABLE;
Disable   := State.eProgress;
END_METHOD

METHOD Reset : E_PROGRESS
VAR_INPUT
END_VAR
Ctrl.eCmd := AXIS_RESET;
Reset     := State.eProgress;
END_METHOD

METHOD Home : E_PROGRESS
VAR_INPUT
END_VAR
Ctrl.eCmd := AXIS_HOME;
Home      := State.eProgress;
END_METHOD

METHOD MoveAbsolute : E_PROGRESS
VAR_INPUT
    lrPosition : LREAL;
    lrVelocity : LREAL;
END_VAR
Ctrl.eCmd             := AXIS_MOVE_ABS;
Data.lrTargetPosition := lrPosition;
Data.lrVelocity       := lrVelocity;
MoveAbsolute          := State.eProgress;
END_METHOD

METHOD MoveRelative : E_PROGRESS
VAR_INPUT
    lrDistance : LREAL;
    lrVelocity : LREAL;
END_VAR
Ctrl.eCmd             := AXIS_MOVE_REL;
Data.lrTargetPosition := lrDistance;
Data.lrVelocity       := lrVelocity;
MoveRelative          := State.eProgress;
END_METHOD

METHOD MoveVelocity : E_PROGRESS
VAR_INPUT
    lrVelocity : LREAL;   // signed
END_VAR
Ctrl.eCmd       := AXIS_MOVE_VELOCITY;
Data.lrVelocity := lrVelocity;
MoveVelocity    := State.eProgress;
END_METHOD

METHOD Jog : E_PROGRESS
VAR_INPUT
    xForward   : BOOL;
    xReverse   : BOOL;
    lrVelocity : LREAL;   // magnitudo
END_VAR
IF    xForward THEN Ctrl.eCmd := AXIS_JOG_POS;
ELSIF xReverse THEN Ctrl.eCmd := AXIS_JOG_NEG;
ELSE               Ctrl.eCmd := AXIS_NULL;
END_IF
Data.lrVelocity := lrVelocity;
Jog             := State.eProgress;
END_METHOD

METHOD MoveFollow : E_PROGRESS
VAR_INPUT
    lrPosition : LREAL;
    lrVelocity : LREAL;
END_VAR
Ctrl.eCmd             := AXIS_MOVE_CSP;
Data.lrTargetPosition := lrPosition;
Data.lrVelocity       := lrVelocity;
MoveFollow            := State.eProgress;
END_METHOD

METHOD Stop : E_PROGRESS
VAR_INPUT
END_VAR
Ctrl.eCmd := AXIS_STOP;
Stop      := State.eProgress;
END_METHOD

PROPERTY Position : LREAL
GET
Position := Info.lrActualPosition;
END_GET
END_PROPERTY

PROPERTY Enabled : BOOL
GET
Enabled := Info.xEnabled;
END_GET
END_PROPERTY

END_FUNCTION_BLOCK

// ---- POUs/SML_Power.TcPOU
(* ============================================================
   SML_Power - CiA402 Drive Power-On / Power-Off Sequencer
   SML v4 - Merged (best of OpenSML_Power + SML_Power/Confa)

   Drives the CiA402 state machine:
     SwitchOnDisabled -> ReadyToSwitchOn -> SwitchedOn -> OperationEnabled

   KEY DESIGN CHOICES (vs original OpenSML):
   - xExecute (edge/level) instead of xEnable:
     After a fault reset the drive returns to Idle and REQUIRES a
     new xExecute pulse.  This prevents automatic re-enable after
     any fault - the operator must consciously re-request power.
   - Single tonTimeout instance with explicit IN management per state.
   - Proper CiA402 Shutdown command on disable (bit3=0, bit0=0).
   - All control bits forced low in error state.

   EMERGENCY STOP:
     xEmergencyStop = TRUE  -> ControlWord bit 2 = 1 -> normal run
     xEmergencyStop = FALSE -> ControlWord bit 2 = 0 -> quick-stop
   Applied every cycle regardless of state.
   ============================================================ *)

FUNCTION_BLOCK SML_Power
VAR_IN_OUT
    Axis : OpenSML_Axis;
END_VAR
VAR_INPUT
    xExecute       : BOOL;           // Level/edge: request drive enable; drop to disable
    xEmergencyStop : BOOL := TRUE;   // TRUE = normal run, FALSE = quick-stop (CiA402 bit 2)
END_VAR
VAR_OUTPUT
    xDone  : BOOL; // Drive in OperationEnabled state, ready for motion FBs
    xError : BOOL; // Fault present or power-up sequence timed out
    eProgress : E_PROGRESS; // Level A: unified progress (projection of iState)
END_VAR
VAR
    iState     : INT;
    tonTimeout : TON;
    tTimeOut   : TIME := T#500MS; // Max time allowed per CiA402 state transition
END_VAR

// -- Quick-Stop line - written every scan regardless of state --------------
// CiA402 bit 2: 1 = normal, 0 = quick-stop. Active-LOW - never invert here.
Axis.ControlWord.2 := xEmergencyStop;

// -- Single timer instance - IN assigned per state -------------------------
tonTimeout(PT := tTimeOut);

CASE iState OF

    0: // Idle - safe default; wait for execute request
        xDone  := FALSE;
        xError := FALSE;
        tonTimeout.IN := FALSE;
        Axis.ControlWord.0 := FALSE; // Switch On
        Axis.ControlWord.1 := FALSE; // Enable Voltage
        Axis.ControlWord.3 := FALSE; // Enable Operation
        Axis.ControlWord.7 := FALSE; // Fault Reset (pre-clear)
        IF xExecute THEN
            IF Axis.StatusWord.3 THEN
                iState := 10; // Fault active -> reset first
            ELSE
                iState := 20; // No fault -> begin enable sequence
            END_IF
        END_IF

    10: // Fault Reset - pulse bit 7 (rising edge 0->1 clears fault)
        // On success: return to IDLE (not directly to enable).
        // Operator must re-assert xExecute to intentionally re-enable.
        Axis.ControlWord.7 := TRUE;
        tonTimeout.IN := TRUE;
        IF tonTimeout.Q AND NOT Axis.StatusWord.3 THEN
            Axis.ControlWord.7 := FALSE;
            tonTimeout.IN := FALSE;
            iState := 0; // Back to idle - requires deliberate re-enable
        ELSIF tonTimeout.Q THEN
            tonTimeout.IN := FALSE;
            iState := 999; // Drive did not clear fault within timeout
        END_IF

    20: // Enable Voltage - Shutdown command: bit1=1, bit0=0, bit3=0
        // Transitions: SwitchOnDisabled -> ReadyToSwitchOn
        Axis.ControlWord.1 := TRUE;
        tonTimeout.IN := TRUE;
        IF Axis.StatusWord.0 THEN
            // StatusWord bit 0 = Ready to Switch On confirmed
            tonTimeout.IN := FALSE;
            iState := 30;
        ELSIF tonTimeout.Q THEN
            tonTimeout.IN := FALSE;
            iState := 999;
        END_IF

    30: // Switch On - command: bit1=1, bit0=1, bit3=0
        // Transitions: ReadyToSwitchOn -> SwitchedOn
        Axis.ControlWord.0 := TRUE;
        tonTimeout.IN := TRUE;
        IF Axis.StatusWord.0 AND Axis.StatusWord.1 THEN
            // StatusWord bits 0+1 = Switched On confirmed
            tonTimeout.IN := FALSE;
            iState := 40;
        ELSIF tonTimeout.Q THEN
            tonTimeout.IN := FALSE;
            iState := 999;
        END_IF

    40: // Enable Operation - command: bit0=1, bit1=1, bit3=1
        // Transitions: SwitchedOn -> OperationEnabled
        // Freeze target position BEFORE asserting bit3 to prevent a position jump
        Axis.Target_Position := Axis.Position_Actual_Value;
        Axis.ControlWord.3 := TRUE;
        tonTimeout.IN := TRUE;
        IF Axis.StatusWord.0 AND Axis.StatusWord.1 AND Axis.StatusWord.2 THEN
            // OperationEnabled confirmed
            tonTimeout.IN := FALSE;
            iState := 50;
        ELSIF tonTimeout.Q THEN
            tonTimeout.IN := FALSE;
            iState := 999;
        END_IF

    50: // Running - drive in OperationEnabled, accepting setpoints
        xDone := TRUE;
        IF NOT xExecute THEN
            // CiA402 Shutdown: bit3=0 (Disable Operation) + bit0=0 (Switch Off)
            Axis.ControlWord.3 := FALSE;
            Axis.ControlWord.0 := FALSE;
            iState := 0;
        ELSIF Axis.StatusWord.3 THEN
            // Drive fault while running
            iState := 999;
        ELSIF NOT Axis.StatusWord.5 AND xEmergencyStop THEN
            // M3: QuickStopActive (StatusWord bit 5 = 0) but E-stop has been
            // released (xEmergencyStop = TRUE). Depending on quick-stop option
            // code 0x605A the drive may stay in QuickStopActive and NOT auto-
            // recover. Re-run the enable sequence from Switch-On to bring the
            // drive back to OperationEnabled. xDone drops until re-confirmed.
            xDone := FALSE;
            iState := 20;
        END_IF

    999: // Error - latched; reset by dropping xExecute
        tonTimeout.IN := FALSE;
        xDone  := FALSE;
        xError := TRUE;
        Axis.ControlWord.0 := FALSE; // Force low for safety
        Axis.ControlWord.3 := FALSE;
        IF NOT xExecute THEN
            iState := 0;
        END_IF

END_CASE

// -- Level A: unified progress projection (E_PROGRESS) --------------
IF    xError     THEN eProgress := PROGRESS_ERROR;
ELSIF xDone      THEN eProgress := PROGRESS_DONE;      // OperationEnabled (iState 50)
ELSIF iState = 0 THEN eProgress := PROGRESS_INVALID;   // idle
ELSE                  eProgress := PROGRESS_BUSY;       // sequence in progress
END_IF

END_FUNCTION_BLOCK

// ---- POUs/SML_Reset.TcPOU
(* ============================================================
   SML_Reset - CiA402 Fault Reset (standalone FB)
   SML v4 - Merged (from Confa; not present in original OpenSML)

   Pulses ControlWord bit 7 (rising edge 0->1) to clear a drive
   fault independently of the power sequence.

   Use this FB when you need to reset a fault without going through
   the full SML_Power enable sequence, for example to clear a
   non-critical warning while the drive is in a known safe state.

   State machine:
     0 Idle -> 10 Reset pulse -> 20 Done (wait xExecute drop) -> 0
                             -> 999 Error (fault not cleared)
   ============================================================ *)

FUNCTION_BLOCK SML_Reset
VAR_IN_OUT
    Axis : OpenSML_Axis;
END_VAR
VAR_INPUT
    xExecute : BOOL; // Pulse or level: trigger fault reset
END_VAR
VAR_OUTPUT
    xDone  : BOOL; // Fault cleared successfully
    xError : BOOL; // Fault not cleared within timeout
    eProgress : E_PROGRESS; // Level A: unified progress (projection of iState)
END_VAR
VAR
    iState     : INT;
    tonTimeout : TON;
    tTimeOut   : TIME := T#500MS;
END_VAR

CASE iState OF

    0: // Idle - pre-clear bit 7, wait for execute
        Axis.ControlWord.7 := FALSE; // Rising edge requires bit7 to start at 0
        xDone  := FALSE;
        xError := FALSE;
        IF xExecute THEN
            iState := 10;
        END_IF

    10: // Assert Fault Reset bit (rising edge 0->1)
        Axis.ControlWord.7 := TRUE;
        tonTimeout(IN := TRUE, PT := tTimeOut);
        IF tonTimeout.Q AND NOT Axis.StatusWord.3 THEN
            // Fault cleared
            Axis.ControlWord.7 := FALSE;
            xDone := TRUE;
            tonTimeout(IN := FALSE);
            iState := 20;
        ELSIF tonTimeout.Q THEN
            // Persistent fault - hardware intervention required
            Axis.ControlWord.7 := FALSE;
            tonTimeout(IN := FALSE);
            iState := 999;
        END_IF

    20: // Done - hold until xExecute drops (prevents continuous re-reset)
        IF NOT xExecute THEN
            iState := 0;
        END_IF

    999: // Error - fault not cleared; reset by dropping xExecute
        tonTimeout(IN := FALSE);
        Axis.ControlWord.7 := FALSE;
        xError := TRUE;
        IF NOT xExecute THEN
            iState := 0;
        END_IF

END_CASE

// -- Level A: unified progress projection (E_PROGRESS) --------------
IF    xError     THEN eProgress := PROGRESS_ERROR;
ELSIF xDone      THEN eProgress := PROGRESS_DONE;
ELSIF iState = 0 THEN eProgress := PROGRESS_INVALID;
ELSE                  eProgress := PROGRESS_BUSY;
END_IF

END_FUNCTION_BLOCK

// ---- POUs/SML_Home.TcPOU
(* ============================================================
   SML_Home - CiA402 Homing Sequence (mode 6)
   SML v4 - Merged (OpenSML_Home + SML_Home/Confa)

   Prerequisites - configure via SDO or EtherCAT startup params:
     0x6098  Homing Method
     0x6099.01  Speed for limit switch search
     0x6099.02  Speed for index pulse
     0x609A  Homing Acceleration

   The homing offset (0x607C) is written via PDO at runtime
   through diHomeOffset - no SDO access needed.

   CiA402 completion: StatusWord bit 10 (Target Reached) AND
   bit 12 (Home Attained) must both be set.

   State flow:
     0 Idle -> 10 Mode Switch -> 20 Homing -> 30 Done -> 40 Handshake -> 0
                                         -> 999 Error

   Stall watchdog (state 20): if position doesn't change for
   tStallTimeout, the homing sequence is aborted.
   ============================================================ *)

FUNCTION_BLOCK SML_Home
VAR_IN_OUT
    Axis : OpenSML_Axis;
END_VAR
VAR_INPUT
    xEnable        : BOOL;           // Level: FB active; drop to abort
    xExecute       : BOOL;           // Edge/level: start homing
    xReset         : BOOL;           // Pulse: acknowledge error and return to idle
    diHomeOffset   : DINT;           // Home offset [encoder counts] - written to 0x607C
    tStallTimeout  : TIME := T#10S;  // Max time without position change before error
END_VAR
VAR_OUTPUT
    xBusy  : BOOL; // Homing sequence in progress
    xDone  : BOOL; // Homing completed successfully
    xError : BOOL; // Error: fault, stall, timeout, or operator abort
    eProgress : E_PROGRESS; // Level A: unified progress (projection of iState)
END_VAR
VAR
    iState     : INT;
    tonStall   : TON;  // Stall watchdog
    tonMode    : TON;  // Mode-switch timeout guard
    Pos_Old    : DINT; // Previous-cycle position for stall detection
END_VAR

CASE iState OF

    0: // Idle - reset outputs, capture baseline position for stall detection
        xBusy  := FALSE;
        xDone  := FALSE;
        xError := FALSE;
        tonStall.IN := FALSE;
        tonMode.IN  := FALSE;
        Pos_Old := Axis.Position_Actual_Value; // Baseline so state 20 starts correctly

        IF xEnable THEN
            IF xExecute AND Axis.StatusWord.1         // SwitchedOn
                        AND Axis.StatusWord.2         // OperationEnabled
                        AND Axis.Modes_of_operation_display = 6 // Already in Homing mode
                        AND NOT Axis.StatusWord.3 THEN
                iState := 10;

            ELSIF xExecute AND Axis.StatusWord.1
                           AND Axis.Modes_of_operation_display <> 6 THEN
                // Different mode active - drop EnableOperation for mode switch
                Axis.ControlWord.3 := FALSE;
                iState := 10;

            ELSIF xExecute OR Axis.StatusWord.3 THEN
                iState := 999; // Drive not ready or fault present
            END_IF
        END_IF

    10: // Mode Switch - request Homing mode, write offset, re-enable operation
        tonMode(IN := TRUE, PT := T#2S); // Mode switch should be nearly instantaneous
        Axis.ControlWord.4      := FALSE;       // Clear Start Homing bit before arming
        Axis.Modes_of_operation := 6;           // Request Homing mode
        Axis.Home_Offset        := diHomeOffset; // Write offset to 0x607C via PDO

        // Re-enable operation only when drive confirms mode 6 is active
        Axis.ControlWord.3 := (Axis.Modes_of_operation_display = 6);

        IF Axis.StatusWord.3 OR NOT xEnable OR tonMode.Q THEN
            tonMode.IN := FALSE;
            iState := 999;
        ELSIF Axis.StatusWord.2 AND Axis.ControlWord.3 THEN
            // OperationEnabled confirmed in Homing mode
            tonMode.IN := FALSE;
            xBusy := TRUE;
            iState := 20;
        END_IF

    20: // Homing in progress - arm Start Homing, monitor completion and stall
        Axis.ControlWord.4 := TRUE; // Start Homing (bit 4 in HM mode)

        // Stall watchdog: timer runs while position is unchanged from last cycle.
        // Pos_Old updated AFTER timer call so comparison is current-vs-previous.
        tonStall(IN := (Axis.Position_Actual_Value = Pos_Old), PT := tStallTimeout);
        Pos_Old := Axis.Position_Actual_Value;

        IF Axis.StatusWord.3 OR NOT xEnable THEN
            // Drive fault or operator abort
            tonStall.IN := FALSE;
            iState := 999;
        ELSIF tonStall.Q THEN
            // Axis hasn't moved for tStallTimeout -> stalled or misconfigured
            tonStall.IN := FALSE;
            iState := 999;
        ELSIF Axis.StatusWord.10 AND Axis.StatusWord.12 THEN
            // Target Reached (bit 10) AND Home Attained (bit 12) = success
            tonStall.IN := FALSE;
            Axis.ControlWord.4   := FALSE;               // Deassert Start Homing
            Axis.Target_Position := Axis.Position_Actual_Value; // Prevent position jump
            iState := 30;
        END_IF

    30: // Done - hold xDone until xExecute drops
        xDone := TRUE;
        IF NOT xEnable THEN
            iState := 0;
        ELSIF NOT xExecute THEN
            iState := 40; // Wait for handshake before accepting new request
        END_IF

    40: // Handshake - wait here until a new xExecute is asserted or enable drops
        // Prevents bounce if xExecute is held after completion
        IF NOT xEnable THEN
            iState := 0;
        ELSIF xExecute THEN
            // New homing request - go to idle so state 0 evaluates fresh
            iState := 0;
        END_IF

    999: // Error - latched; reset by xReset pulse or dropping xExecute
        tonStall.IN := FALSE;
        tonMode.IN  := FALSE;
        Axis.ControlWord.4 := FALSE; // Deassert Start Homing for safety
        xBusy  := FALSE;
        xError := TRUE;
        IF NOT xExecute OR xReset THEN
            iState := 0;
        END_IF

END_CASE

// -- Level A: unified progress projection (E_PROGRESS) --------------
IF    xError     THEN eProgress := PROGRESS_ERROR;
ELSIF xDone      THEN eProgress := PROGRESS_DONE;
ELSIF iState = 0 THEN eProgress := PROGRESS_INVALID;
ELSE                  eProgress := PROGRESS_BUSY;
END_IF

END_FUNCTION_BLOCK

// ---- POUs/SML_ProfilePosition.TcPOU
(* ============================================================
   SML_ProfilePosition - CiA402 Profile Position Mode (PP, mode 1)
   SML v4 - Merged (OpenSML_ProfilePosition + SML_ProfilePosition/Confa)

   Profile Acceleration and Deceleration are passed per-call and
   written to Axis.Profile_Acceleration / Axis.Profile_Deceleration
   (0x6083 / 0x6084) via PDO - no SDO access required.

   CiA402 PP setpoint protocol (implemented via states 10->20->30->40):
     1. Write Target_Position, Profile_Velocity, Accel, Decel
     2. Set ControlWord bit 4 (New Setpoint) = 1
     3. Wait StatusWord bit 12 (Setpoint Acknowledge) = 1
     4. Clear ControlWord bit 4 = 0
     5. Wait StatusWord bit 10 (Target Reached) = 1

   States:
     0   Idle - wait for enable + execute
     10  Mode Switch - switch to PP mode 1
     20  Setpoint active - wait for acknowledge / target / error
     30  Acknowledged - wait for target reached or new execute
     40  Target reached - hold xDone until execute drops
     999 Error - hold position; reset by xReset or NOT xEnable
   ============================================================ *)

FUNCTION_BLOCK SML_ProfilePosition
VAR_IN_OUT
    Axis : OpenSML_Axis;
END_VAR
VAR_INPUT
    xEnable                : BOOL;   // Level: keep FB active
    xExecute               : BOOL;   // Trigger: start move (hold for duration)
    xContinueMove          : BOOL;   // Blend: no deceleration between consecutive moves (bit 5)
    xRelativeMode          : BOOL;   // FALSE = absolute, TRUE = relative (bit 6)
    xReset                 : BOOL;   // Pulse: acknowledge error
    diTargetPosition       : DINT;   // Target [encoder counts, raw drive units]
    udiProfileVelocity     : UDINT;  // Move speed [drive velocity units]; must be > 0
    udiProfileAcceleration : UDINT;  // Acceleration [drive accel units]
    udiProfileDeceleration : UDINT;  // Deceleration [drive accel units]
END_VAR
VAR_OUTPUT
    xDone   : BOOL; // Target position reached (bit 10 set, no following error)
    xBusy   : BOOL; // Setpoint acknowledged (bit 12), motion in progress
    xMoving : BOOL; // Axis velocity <> 0 (StatusWord bit 14 = 0 on many drives)
    xError  : BOOL; // Fault (bit 3) or following error (bit 13)
    eProgress : E_PROGRESS; // Level A: unified progress (projection of iState)
END_VAR
VAR
    iState : INT;
END_VAR

// -- Continuous outputs (updated every cycle while in PP mode) -------------
// xBusy: setpoint acknowledged AND target not yet reached
IF xEnable AND Axis.Modes_of_operation_display = 1 THEN
    xBusy := (iState > 0 AND iState < 999)
             AND Axis.StatusWord.12    // Setpoint Acknowledge
             AND NOT Axis.StatusWord.10; // NOT Target Reached
END_IF

// xMoving: bit 14 = standstill flag (0 = moving) - drive-dependent
xMoving := NOT Axis.StatusWord.14;

// -- Write ramp parameters only when commanded -----------------------------
IF xExecute THEN
    Axis.Profile_Acceleration := udiProfileAcceleration;
    Axis.Profile_Deceleration := udiProfileDeceleration;
END_IF

CASE iState OF

    0: // Idle
        xDone  := FALSE;
        xError := FALSE;

        IF xEnable THEN
            IF xExecute AND Axis.StatusWord.1 AND NOT Axis.StatusWord.3 THEN
                // Drive is at least SwitchedOn and no fault - attempt move
                Axis.ControlWord.5    := xContinueMove;
                Axis.ControlWord.6    := xRelativeMode;
                Axis.Profile_Velocity := udiProfileVelocity;
                Axis.Target_Position  := diTargetPosition;
                iState := 10;
            ELSIF xExecute OR Axis.StatusWord.3 THEN
                iState := 999;
            END_IF
        END_IF

    10: // Mode Switch - request PP (mode 1), re-enable operation when confirmed
        Axis.Modes_of_operation := 1;
        Axis.ControlWord.3 := (Axis.Modes_of_operation_display = 1);

        IF Axis.StatusWord.3 OR NOT xEnable THEN
            iState := 999;
        ELSIF Axis.StatusWord.2 AND Axis.Modes_of_operation_display = 1 THEN
            // OperationEnabled in PP mode -> trigger new setpoint (rising edge on bit 4)
            Axis.ControlWord.4 := TRUE;
            iState := 20;
        END_IF

    20: // Active - setpoint sent, waiting for acknowledge/target/error
        IF Axis.StatusWord.13 OR Axis.StatusWord.3 OR NOT xEnable THEN
            // Following error, fault, or operator cancel
            iState := 999;
        ELSIF Axis.StatusWord.10 THEN
            // Target Reached (bit 10) - move complete
            xDone := TRUE;
            Axis.ControlWord.4 := FALSE;
            iState := 40;
        ELSIF Axis.StatusWord.12 AND NOT xExecute THEN
            // Setpoint acknowledged but xExecute already dropped
            // -> clear bit 4 and move to ready-for-next state
            Axis.ControlWord.4 := FALSE;
            iState := 30;
        ELSIF NOT Axis.StatusWord.12 AND NOT Axis.StatusWord.10 AND NOT xExecute THEN
            // Neither acknowledged nor reached, execute dropped -> clean exit
            Axis.ControlWord.4 := FALSE;
            iState := 0;
        END_IF

    30: // Acknowledged - moving toward target; accept next execute or wait
        IF Axis.StatusWord.13 OR Axis.StatusWord.3 OR NOT xEnable THEN
            iState := 999;
        ELSIF Axis.StatusWord.10 THEN
            xDone := TRUE;
            Axis.ControlWord.4 := FALSE;
            iState := 40;
        ELSIF xExecute AND Axis.StatusWord.1 AND NOT Axis.StatusWord.3 THEN
            // New move requested - queue it
            Axis.ControlWord.5    := xContinueMove;
            Axis.ControlWord.6    := xRelativeMode;
            Axis.Profile_Velocity := udiProfileVelocity;
            Axis.Target_Position  := diTargetPosition;
            iState := 10;
        END_IF

    40: // Target reached - hold xDone until execute or enable drops
        IF NOT xEnable OR NOT xExecute THEN
            xDone  := FALSE;
            iState := 0;
        END_IF

    999: // Error - hold current position; reset by xReset or dropping xEnable
        Axis.Profile_Velocity := 0;
        // SAFETY: hold current position, never write 0 (that commands a move to origin)
        Axis.Target_Position  := Axis.Position_Actual_Value;
        Axis.ControlWord.4    := FALSE;
        xError := TRUE;
        IF NOT xEnable OR xReset THEN
            xError := FALSE;
            iState := 0;
        END_IF

END_CASE

// -- Level A: unified progress projection (E_PROGRESS) --------------
IF    xError     THEN eProgress := PROGRESS_ERROR;
ELSIF xDone      THEN eProgress := PROGRESS_DONE;
ELSIF iState = 0 THEN eProgress := PROGRESS_INVALID;
ELSE                  eProgress := PROGRESS_BUSY;
END_IF

END_FUNCTION_BLOCK

// ---- POUs/SML_ProfileVelocity.TcPOU
(* ============================================================
   SML_ProfileVelocity - CiA402 Profile Velocity Mode (PV, mode 3)
   SML v4 - Merged (OpenSML_ProfileVelocity + SML_ProfileVelocity/Confa)

   Profile Acceleration and Deceleration per-call via PDO.
   Drive ramps to diTargetVelocity using its internal planner.
   Signed velocity: positive = forward, negative = reverse, 0 = stop.

   Both following error (bit 13) and fault (bit 3) are monitored
   in the active state.
   ============================================================ *)

FUNCTION_BLOCK SML_ProfileVelocity
VAR_IN_OUT
    Axis : OpenSML_Axis;
END_VAR
VAR_INPUT
    xEnable                : BOOL;   // Level: keep FB active
    xExecute               : BOOL;   // Level/edge: activate velocity mode
    xReset                 : BOOL;   // Pulse: acknowledge error
    diTargetVelocity       : DINT;   // Target velocity [drive units]; signed; 0 = decelerate to stop
    udiProfileAcceleration : UDINT;  // Acceleration [drive accel units]
    udiProfileDeceleration : UDINT;  // Deceleration [drive accel units]
END_VAR
VAR_OUTPUT
    xMoving     : BOOL; // TRUE when axis velocity <> 0 in either direction
    xAtVelocity : BOOL; // TRUE when drive reports target velocity reached (bit 10)
    xError      : BOOL; // Fault or following error
    eProgress   : E_PROGRESS; // Level A: unified progress (projection of iState)
END_VAR
VAR
    iState : INT;
END_VAR

// -- xMoving: detect motion in BOTH forward and reverse --------------------
// ABS() is required - Target_Velocity < 0 during reverse would miss a plain > 0 check
xMoving := NOT Axis.StatusWord.14         // Standstill bit = 0 means moving
           AND ABS(Axis.Target_Velocity) > 0
           AND Axis.Modes_of_operation = 3
           AND Axis.ControlWord.3;

// -- Write ramp params only when a velocity command is active --------------
IF xExecute THEN
    Axis.Profile_Acceleration := udiProfileAcceleration;
    Axis.Profile_Deceleration := udiProfileDeceleration;
END_IF

CASE iState OF

    0: // Idle
        xError      := FALSE;
        xAtVelocity := FALSE;

        IF xEnable THEN
            IF xExecute AND Axis.StatusWord.1          // SwitchedOn
                        AND Axis.StatusWord.2           // Already OperationEnabled
                        AND Axis.Modes_of_operation_display = 3 // Already in PV mode
                        AND NOT Axis.StatusWord.3 THEN
                // M4: fast path - already enabled in PV mode, skip the
                // disable/enable cycle that v3 forced on every start.
                Axis.Target_Velocity := 0;
                iState := 20;
            ELSIF xExecute AND Axis.StatusWord.1       // SwitchedOn
                        AND NOT Axis.StatusWord.2       // Not yet OperationEnabled (needs mode switch)
                        AND NOT Axis.StatusWord.3 THEN
                iState := 10;
            ELSIF xExecute AND Axis.StatusWord.2 THEN
                // OperationEnabled but wrong mode - drop bit3 for switch
                Axis.ControlWord.3 := FALSE;
                // State stays 0: StatusWord.2 drops next cycle, mode-switch branch fires
            ELSIF xExecute OR Axis.StatusWord.3 THEN
                iState := 999;
            END_IF
        END_IF

    10: // Mode Switch - request PV (mode 3)
        Axis.Modes_of_operation := 3;
        Axis.ControlWord.3 := (Axis.Modes_of_operation_display = 3);

        IF Axis.StatusWord.3 OR NOT xEnable THEN
            iState := 999;
        ELSIF Axis.StatusWord.2 AND Axis.ControlWord.3 THEN
            // OperationEnabled in PV mode - zero velocity on entry
            Axis.Target_Velocity := 0;
            iState := 20;
        END_IF

    20: // Active - write velocity every cycle
        IF Axis.Modes_of_operation_display = 3 THEN
            Axis.Target_Velocity := diTargetVelocity;
            xAtVelocity := Axis.StatusWord.10; // "Target velocity reached" in PV mode

            IF Axis.StatusWord.3 THEN
                // Drive fault
                Axis.Target_Velocity := 0;
                iState := 999;
            ELSIF Axis.StatusWord.13 THEN
                // Following error
                Axis.Target_Velocity := 0;
                iState := 999;
            ELSIF NOT xEnable THEN
                // Normal stop: write 0 -> drive decelerates using Profile_Deceleration
                Axis.Target_Velocity := 0;
                iState := 0;
            END_IF
        ELSE
            // Drive changed mode unexpectedly
            Axis.Target_Velocity := 0;
            iState := 0;
        END_IF

    999: // Error
        Axis.Target_Velocity  := 0;
        Axis.Profile_Velocity := 0; // Also clear PP speed register
        xError      := TRUE;
        xAtVelocity := FALSE;
        IF NOT xExecute OR xReset THEN
            xError := FALSE;
            iState := 0;
        END_IF

END_CASE

// -- Level A: unified progress projection (E_PROGRESS) --------------
// Continuous mode: "DONE" = target velocity reached (steady state).
IF    xError       THEN eProgress := PROGRESS_ERROR;
ELSIF xAtVelocity  THEN eProgress := PROGRESS_DONE;
ELSIF iState = 0   THEN eProgress := PROGRESS_INVALID;
ELSE                    eProgress := PROGRESS_BUSY;
END_IF

END_FUNCTION_BLOCK

// ---- POUs/SML_ProfileVelocity_Jog.TcPOU
(* ============================================================
   SML_ProfileVelocity_Jog - Dedicated Jog FB (PV mode 3)
   SML v4 - Merged (from Confa; improved state machine)

   Provides separate hold-to-run forward/reverse inputs.
   FB stays in state 20 as long as xEnable is TRUE, avoiding
   a mode-switch cycle every time the jog button is released.
   Returns to idle only on xEnable drop.

   Velocity is always derived from ABS(diProfileVelocity) and
   negated for reverse - eliminates double-negation risk.
   ============================================================ *)

FUNCTION_BLOCK SML_ProfileVelocity_Jog
VAR_IN_OUT
    Axis : OpenSML_Axis;
END_VAR
VAR_INPUT
    xEnable                : BOOL;   // Level: keep FB active
    xExecute_Jog_F         : BOOL;   // Hold: jog forward (positive velocity)
    xExecute_Jog_R         : BOOL;   // Hold: jog reverse (negative velocity)
    xReset                 : BOOL;   // Pulse: acknowledge error
    diProfileVelocity      : DINT;   // Speed magnitude [drive units]; must be > 0
    udiProfileAcceleration : UDINT;  // Acceleration [drive accel units]
    udiProfileDeceleration : UDINT;  // Deceleration [drive accel units]
END_VAR
VAR_OUTPUT
    xMoving : BOOL; // TRUE when axis velocity <> 0 in either direction
    xError  : BOOL; // Drive fault detected
    eProgress : E_PROGRESS; // Level A: unified progress (projection of iState)
END_VAR
VAR
    xAnyJog : BOOL; // Internal: TRUE if either direction is active
    iState  : INT;
END_VAR

// -- Internal execute: jog active if either direction AND enabled ----------
xAnyJog := (xExecute_Jog_F OR xExecute_Jog_R) AND xEnable;

// -- xMoving: detect motion in both directions -----------------------------
xMoving := NOT Axis.StatusWord.14
           AND ABS(Axis.Target_Velocity) > 0
           AND Axis.Modes_of_operation = 3
           AND Axis.ControlWord.3;

// -- Write ramp params only when jogging -----------------------------------
IF xAnyJog THEN
    Axis.Profile_Acceleration := udiProfileAcceleration;
    Axis.Profile_Deceleration := udiProfileDeceleration;
END_IF

CASE iState OF

    0: // Idle
        xError := FALSE;
        IF xEnable THEN
            IF xAnyJog AND Axis.StatusWord.1 AND NOT Axis.StatusWord.3 THEN
                IF Axis.StatusWord.2 AND Axis.Modes_of_operation_display = 3 THEN
                    // M4: fast path - already enabled in PV mode, jog immediately.
                    Axis.Target_Velocity := 0;
                    iState := 20;
                ELSIF NOT Axis.StatusWord.2 THEN
                    iState := 10; // SwitchedOn but not OperationEnabled -> mode switch
                ELSE
                    // OperationEnabled but wrong mode - drop bit3 to allow mode switch
                    Axis.ControlWord.3 := FALSE;
                    // State stays 0; StatusWord.2 drops next cycle -> mode-switch branch fires
                END_IF
            ELSIF xAnyJog OR Axis.StatusWord.3 THEN
                iState := 999;
            END_IF
        END_IF

    10: // Mode Switch - request PV (mode 3)
        Axis.Modes_of_operation := 3;
        Axis.ControlWord.3 := (Axis.Modes_of_operation_display = 3);

        IF Axis.StatusWord.3 OR NOT xEnable THEN
            iState := 999;
        ELSIF Axis.StatusWord.2 AND Axis.ControlWord.3 THEN
            Axis.Target_Velocity := 0; // Zero on entry
            iState := 20;
        END_IF

    20: // Jog active - stays here while xEnable is TRUE
        IF Axis.Modes_of_operation_display = 3 THEN
            IF Axis.StatusWord.3 OR NOT xEnable THEN
                // Fault or operator disable
                Axis.Target_Velocity := 0;
                iState := 999;

            ELSIF xExecute_Jog_F AND NOT xExecute_Jog_R THEN
                // Forward: always positive (ABS prevents sign surprises)
                Axis.Target_Velocity := ABS(diProfileVelocity);

            ELSIF xExecute_Jog_R AND NOT xExecute_Jog_F THEN
                // Reverse: negate magnitude
                Axis.Target_Velocity := -ABS(diProfileVelocity);

            ELSE
                // No jog or both simultaneously -> decelerate and hold in mode
                // STAY in state 20: no mode-switch latency on next jog press
                Axis.Target_Velocity := 0;
            END_IF
        ELSE
            // Drive changed mode unexpectedly
            Axis.Target_Velocity := 0;
            iState := 0;
        END_IF

    999: // Error
        Axis.Target_Velocity  := 0;
        Axis.Profile_Velocity := 0;
        xError := TRUE;
        IF NOT xAnyJog OR xReset THEN
            xError := FALSE;
            iState := 0;
        END_IF

END_CASE

// -- Level A: unified progress projection (E_PROGRESS) --------------
// Jog is a held continuous motion: no discrete "DONE".
IF    xError     THEN eProgress := PROGRESS_ERROR;
ELSIF iState = 0 THEN eProgress := PROGRESS_INVALID;
ELSE                  eProgress := PROGRESS_BUSY;      // jog in progress
END_IF

END_FUNCTION_BLOCK

// ---- POUs/SML_Stop.TcPOU
(* ============================================================
   SML_Stop - CiA402 Halt (software controlled stop)
   SML v4 - Merged (OpenSML_Stop + Confa SML_Stop + xStopped output)

   Sets ControlWord bit 8 (Halt):
   - xStop = TRUE : drive decelerates to zero using Profile_Deceleration;
     drive stays in OperationEnabled and holds position
   - xStop = FALSE: motion FBs can resume commanding the axis

   This is a SOFT stop - the axis decelerates under control.
   For an emergency HARD stop use xEmergencyStop = FALSE via
   SML_Power (sets ControlWord bit 2 = 0 -> quick-stop deceleration).

   xStopped: TRUE when Halt is active AND the drive reports that
   velocity has reached zero.  StatusWord bit 10 meaning is
   operating-mode dependent - verify against your drive datasheet.
   ============================================================ *)

FUNCTION_BLOCK SML_Stop
VAR_IN_OUT
    Axis : OpenSML_Axis;
END_VAR
VAR_INPUT
    xStop : BOOL; // TRUE = activate Halt; FALSE = release Halt
END_VAR
VAR_OUTPUT
    xStopped : BOOL; // TRUE when Halt active and drive reports standstill
    eProgress : E_PROGRESS; // Level A: unified progress
END_VAR

// -- Halt bit (ControlWord bit 8) - every cycle ----------------------------
Axis.ControlWord.8 := xStop;

// -- Standstill confirmation -----------------------------------------------
// Only meaningful while xStop is active.
// Bit 10 = "Target Reached" in PP mode, "At Velocity" in PV mode,
// and "Drive Halted" / "Speed Zero" on many drives in Halt condition.
xStopped := xStop AND Axis.StatusWord.10;

// -- Level A: unified progress projection (E_PROGRESS) --------------
IF    NOT xStop  THEN eProgress := PROGRESS_INVALID;
ELSIF xStopped   THEN eProgress := PROGRESS_DONE;
ELSE                  eProgress := PROGRESS_BUSY;   // decelerating
END_IF

END_FUNCTION_BLOCK

// ---- POUs/SML_Diagnostics.TcPOU
(* ============================================================
   SML_Diagnostics - Aggregated Runtime Diagnostics
   SML v4 - New in v4

   PURPOSE
   Turns scattered status bits and per-FB error flags into a single,
   clear diagnostic picture for the operator / HMI:
     - one prioritized current condition (DiagCode + DiagText)
     - a LATCHED first-cause (FirstFaultCode + FirstFaultText) so the
       root cause survives even after follow-on faults pile up
     - explicit fault vs warning classification
     - drive Error_Code (0x603F) and Following_Error (0x60F4) surfaced
     - a cumulative fault event counter for maintenance

   WHY A FIRST-FAULT LATCH?
   When a drive faults, many bits trip at once (fault + following error +
   quick-stop). The operator needs to know WHICH came first. DiagCode
   shows the live highest-priority condition; FirstFaultCode freezes the
   first fault seen until xReset.

   PRIORITY (highest first) for the live DiagCode:
     1 Drive fault (with/without Error_Code)   2 Quick-stop active
     3 Following error                          4 Power FB error
     5 Home error    6 Move error   7 Velocity error
     8 Jog error     9 Touch-probe error       10 OTG error
    11 Internal limit (warning)                12 Drive warning
       otherwise OK

   INTEGRATION
   Call once per cycle. Wire the per-FB xError outputs from FB_SML
   (or your own application) into the xXxxError inputs. Axis gives the
   drive-level bits directly. Reset the latch with a pulse on xReset.

   NOTE: DiagText carries only the category. The numeric drive code is
   in DriveErrorCode (compose "Drive error " + code on the HMI if needed)
   - this keeps the FB free of string-library dependencies.
   ============================================================ *)

FUNCTION_BLOCK SML_Diagnostics
VAR_IN_OUT
    Axis : OpenSML_Axis;
END_VAR
VAR_INPUT
    xReset           : BOOL;   // Pulse: clear the latched first-fault (and acknowledge)
    xResetCount      : BOOL;   // Pulse: clear the cumulative FaultCount

    // -- Aggregated per-FB error flags (wire from FB_SML / application) --
    xPowerError      : BOOL;
    xHomeError       : BOOL;
    xMoveError       : BOOL;   // ProfilePosition (MoveAbs + MoveHome)
    xVelError        : BOOL;
    xJogError        : BOOL;
    xTouchProbeError : BOOL;
    xOtgError        : BOOL;   // FB_S7RTT_OTG constraint error (CSP/OTG paths)
END_VAR
VAR_OUTPUT
    // -- Live condition ----------------------------------------
    DiagCode       : SML_DiagCode;  // Highest-priority active condition this cycle
    DiagText       : STRING(80);    // Human-readable text for DiagCode
    xActiveFault   : BOOL;          // TRUE while any fault condition is present
    xActiveWarning : BOOL;          // TRUE while a warning (no fault) is present

    // -- Latched first cause -----------------------------------
    FirstFaultCode : SML_DiagCode;  // First fault seen since last xReset
    FirstFaultText : STRING(80);    // Text of the first fault

    // -- Drive detail (always live) ----------------------------
    DriveErrorCode : UINT;          // 0x603F raw drive error number (0 = none)
    FollowingError : DINT;          // 0x60F4 following error [encoder counts]

    // -- Maintenance -------------------------------------------
    FaultCount     : UINT;          // Cumulative count of fault events (rising edges)
END_VAR
VAR
    _quickStop : BOOL;  // QuickStopActive decoded from StatusWord
    _prevFault : BOOL;  // Edge detect for FaultCount / first-fault latch
END_VAR

// -- Always-live drive detail -----------------------------------------------
DriveErrorCode := Axis.Error_Code;
FollowingError := Axis.Following_Error_Actual_Value;

// QuickStopActive (CiA402 Table 28): bits 0,1,2 = 1 AND bit 5 = 0
_quickStop := Axis.StatusWord.0 AND Axis.StatusWord.1 AND Axis.StatusWord.2
              AND NOT Axis.StatusWord.5;

// -- Determine the live condition by priority -------------------------------
IF Axis.StatusWord.3 THEN
    // Drive fault - distinguish coded vs uncoded
    IF Axis.Error_Code > 0 THEN
        DiagCode := DIAG_DRIVE_ERRORCODE;
        DiagText := 'Drive fault - see DriveErrorCode (0x603F)';
    ELSE
        DiagCode := DIAG_DRIVE_FAULT;
        DiagText := 'Drive fault - StatusWord bit 3';
    END_IF

ELSIF _quickStop THEN
    DiagCode := DIAG_QUICK_STOP;
    DiagText := 'Quick-stop active - E-stop / ControlWord bit 2';

ELSIF Axis.StatusWord.13 THEN
    DiagCode := DIAG_FOLLOWING_ERROR;
    DiagText := 'Following error - StatusWord bit 13';

ELSIF xPowerError THEN
    DiagCode := DIAG_POWER_ERROR;
    DiagText := 'Power sequence error - SML_Power timed out';

ELSIF xHomeError THEN
    DiagCode := DIAG_HOME_ERROR;
    DiagText := 'Homing error - stall / timeout / abort';

ELSIF xMoveError THEN
    DiagCode := DIAG_MOVE_ERROR;
    DiagText := 'Position move error - ProfilePosition';

ELSIF xVelError THEN
    DiagCode := DIAG_VEL_ERROR;
    DiagText := 'Velocity move error - ProfileVelocity';

ELSIF xJogError THEN
    DiagCode := DIAG_JOG_ERROR;
    DiagText := 'Jog error - ProfileVelocity_Jog';

ELSIF xTouchProbeError THEN
    DiagCode := DIAG_TOUCHPROBE_ERROR;
    DiagText := 'Touch-probe error - capture/enable timeout';

ELSIF xOtgError THEN
    DiagCode := DIAG_OTG_ERROR;
    DiagText := 'OTG error - invalid limits or cycle time';

ELSIF Axis.StatusWord.11 THEN
    DiagCode := DIAG_INTERNAL_LIMIT;
    DiagText := 'Warning - internal limit active (StatusWord bit 11)';

ELSIF Axis.StatusWord.7 THEN
    DiagCode := DIAG_WARNING;
    DiagText := 'Warning - drive warning (StatusWord bit 7)';

ELSE
    DiagCode := DIAG_OK;
    DiagText := 'OK';
END_IF

// -- Classify (codes >= DIAG_DRIVE_FAULT (10) are faults; 1..9 warnings) ----
xActiveFault   := (DiagCode >= DIAG_DRIVE_FAULT);
xActiveWarning := (DiagCode >= DIAG_WARNING) AND (DiagCode < DIAG_DRIVE_FAULT);

// -- First-fault latch + fault event counter (rising edge of any fault) -----
IF xActiveFault AND NOT _prevFault THEN
    FaultCount := FaultCount + 1;
    IF FirstFaultCode = DIAG_OK THEN
        FirstFaultCode := DiagCode;
        FirstFaultText := DiagText;
    END_IF
END_IF
_prevFault := xActiveFault;

// -- Acknowledge / reset ----------------------------------------------------
IF xReset THEN
    FirstFaultCode := DIAG_OK;
    FirstFaultText := 'OK';
END_IF
IF xResetCount THEN
    FaultCount := 0;
END_IF

END_FUNCTION_BLOCK

// ---- POUs/SML_Status.TcPOU
(* ============================================================
   SML_Status - CiA402 StatusWord Decoder + Position/Speed Readout
   SML v4 - Merged (from Confa; not in original OpenSML)

   Decodes the CiA402 state machine and all relevant status bits
   into named BOOL flags.  Useful for HMI display, interlock
   logic, and diagnostics.

   CiA402 state machine (Table 28), identified by bits 6,5,3,2,1,0:
     NotReadyToSwitchOn   : bits = x0 0000  (bit6=0)
     SwitchOnDisabled     : bits = x1 0000  (bit6=1)
     ReadyToSwitchOn      : bits = 01 0001  (bit5=1, bit0=1)
     SwitchedOn           : bits = 01 0011  (bit5=1, bits0-1=1)
     OperationEnabled     : bits = 01 0111  (bit5=1, bits0-2=1)
     QuickStopActive      : bits = 00 0111  (bit5=0, bits0-2=1)
     FaultReactionActive  : bits = x0 1111  (bit3=1, bits0-2=1)
     Fault                : bits = x0 1000  (bit3=1, bits0-2=0)

   DRIVE-SPECIFIC NOTES:
   - Status_Homed reads Digital_Inputs bit 0 (0x60FD).
     Requires the drive configured to set DI0 when homing completes.
     If unsupported, use HomeDone from FB_SML instead.
   - STANDSTILL_THRESHOLD is in drive velocity units.
     Adjust to match your drive's velocity scaling.
   ============================================================ *)

FUNCTION_BLOCK SML_Status
VAR_IN_OUT
    Axis : OpenSML_Axis;
END_VAR
VAR_INPUT
    xEnable : BOOL; // Level: enable decoding
END_VAR
VAR_OUTPUT
    // -- CiA402 state machine ----------------------------------
    Status_NotReadyToSwitchOn  : BOOL;
    Status_SwitchOnDisabled    : BOOL;
    Status_ReadyToSwitchOn     : BOOL;
    Status_SwitchedOn          : BOOL;
    Status_OperationEnabled    : BOOL;
    Status_QuickStopActive     : BOOL;
    Status_FaultReactionActive : BOOL;
    Status_Fault               : BOOL;
    // -- General status ----------------------------------------
    Status_Warning             : BOOL; // Non-fatal (bit 7)
    Status_TargetReached       : BOOL; // Mode-dependent (bit 10)
    Status_Halted              : BOOL; // Halt active + standstill confirmed
    Status_VoltageEnabled      : BOOL; // DC bus present (bit 4)
    Status_InternalLimit       : BOOL; // Software limit active (bit 11)
    // -- Operating mode ----------------------------------------
    Status_ProfilePositionMode : BOOL; // Active mode = PP (1)
    Status_ProfileVelocityMode : BOOL; // Active mode = PV (3)
    Status_VelocityMode        : BOOL; // Active mode = Velocity (2, legacy)
    Status_TorqueProfileMode   : BOOL; // Active mode = Torque (4)
    Status_HomingMode          : BOOL; // Active mode = Homing (6)
    Status_SyncPositionMode    : BOOL; // Active mode = CSP (8)
    Status_SyncVelocityMode    : BOOL; // Active mode = CSV (9)
    // -- Motion ------------------------------------------------
    Status_Moving              : BOOL; // ABS(velocity) > threshold
    Status_StandStill          : BOOL; // ABS(velocity) <= threshold
    Status_Homed               : BOOL; // Drive DI0 = homed (drive-specific)
    // -- Error -------------------------------------------------
    StatusErr                  : BOOL; // Error_Code PDO is non-zero
    ErrId                      : UINT; // Drive error number (0x603F)
    // -- Actual values -----------------------------------------
    ActPosition                : DINT; // [encoder counts]
    ActSpeed                   : DINT; // [drive velocity units]
    ActTorque                  : INT;  // [0.1 % of rated]
    FollowingError             : DINT; // [encoder counts]
END_VAR

VAR CONSTANT
    STANDSTILL_THRESHOLD : DINT := 10; // Velocity units below which axis is "at rest"
END_VAR

IF NOT xEnable THEN RETURN; END_IF

// -- Error code ------------------------------------------------------------
StatusErr := Axis.Error_Code > 0;
ErrId     := Axis.Error_Code;

// -- CiA402 state machine decode ------------------------------------------
Status_NotReadyToSwitchOn :=
    NOT Axis.StatusWord.0 AND NOT Axis.StatusWord.1 AND NOT Axis.StatusWord.2
    AND NOT Axis.StatusWord.3 AND NOT Axis.StatusWord.6;

Status_SwitchOnDisabled :=
    NOT Axis.StatusWord.0 AND NOT Axis.StatusWord.1 AND NOT Axis.StatusWord.2
    AND NOT Axis.StatusWord.3 AND Axis.StatusWord.6;

Status_ReadyToSwitchOn :=
    Axis.StatusWord.0 AND NOT Axis.StatusWord.1 AND NOT Axis.StatusWord.2
    AND NOT Axis.StatusWord.3 AND Axis.StatusWord.5 AND NOT Axis.StatusWord.6;

Status_SwitchedOn :=
    Axis.StatusWord.0 AND Axis.StatusWord.1 AND NOT Axis.StatusWord.2
    AND NOT Axis.StatusWord.3 AND Axis.StatusWord.5 AND NOT Axis.StatusWord.6;

Status_OperationEnabled :=
    Axis.StatusWord.0 AND Axis.StatusWord.1 AND Axis.StatusWord.2
    AND NOT Axis.StatusWord.3 AND Axis.StatusWord.5 AND NOT Axis.StatusWord.6;

Status_QuickStopActive :=
    Axis.StatusWord.0 AND Axis.StatusWord.1 AND Axis.StatusWord.2
    AND NOT Axis.StatusWord.3 AND NOT Axis.StatusWord.5 AND NOT Axis.StatusWord.6;

Status_FaultReactionActive :=
    Axis.StatusWord.0 AND Axis.StatusWord.1 AND Axis.StatusWord.2
    AND Axis.StatusWord.3 AND NOT Axis.StatusWord.6;

Status_Fault :=
    NOT Axis.StatusWord.0 AND NOT Axis.StatusWord.1 AND NOT Axis.StatusWord.2
    AND Axis.StatusWord.3 AND NOT Axis.StatusWord.6;

// -- General status bits ---------------------------------------------------
Status_Warning        := Axis.StatusWord.7;   // Non-fatal warning
Status_TargetReached  := Axis.StatusWord.10;  // Move complete / at velocity (mode-dependent)
Status_InternalLimit  := Axis.StatusWord.11;  // Software limit reached
Status_VoltageEnabled := Axis.StatusWord.4;   // DC bus energized
Status_Halted         := Axis.ControlWord.8 AND Axis.StatusWord.10;

// -- Operating mode --------------------------------------------------------
Status_ProfilePositionMode := (Axis.Modes_of_operation_display = 1);
Status_VelocityMode        := (Axis.Modes_of_operation_display = 2);
Status_ProfileVelocityMode := (Axis.Modes_of_operation_display = 3);
Status_TorqueProfileMode   := (Axis.Modes_of_operation_display = 4);
Status_HomingMode          := (Axis.Modes_of_operation_display = 6);
Status_SyncPositionMode    := (Axis.Modes_of_operation_display = 8);
Status_SyncVelocityMode    := (Axis.Modes_of_operation_display = 9);

// -- Motion detection - consistent threshold (no dead zone) ---------------
Status_Moving     := ABS(Axis.Velocity_Actual_Value) > STANDSTILL_THRESHOLD;
Status_StandStill := ABS(Axis.Velocity_Actual_Value) <= STANDSTILL_THRESHOLD;

// -- Actual values ---------------------------------------------------------
ActPosition    := Axis.Position_Actual_Value;
ActSpeed       := Axis.Velocity_Actual_Value;
ActTorque      := Axis.Torque_Actual_Value;
FollowingError := Axis.Following_Error_Actual_Value;

// -- Homed flag (drive-specific - requires DI0 configured for homed status) -
Status_Homed := Axis.Digital_Inputs.0;

END_FUNCTION_BLOCK

// ---- POUs/SML_TouchProbe.TcPOU
(* ============================================================
   SML_TouchProbe - CiA402 Touch Probe (high-speed position latch)
   SML v4 - Merged (from Confa; added capture timeout)

   Objects used:
     0x60B8  TouchProbe_ControlWord  (output)
     0x60B9  TouchProbe_StatusWord   (input)
     0x60BA  TouchProbe_Rising_Value  [encoder counts] (input)
     0x60BB  TouchProbe_Falling_Value [encoder counts] (input)

   ControlWord 0x60B8:
     Bit 0  Enable Touch Probe 1
     Bit 1  Capture mode (0=single, 1=continuous)
     Bit 2  Trigger source (0=DI13, 1=encoder Z-pulse)
     Bit 4  Enable rising-edge capture -> 0x60BA
     Bit 5  Enable falling-edge capture -> 0x60BB

   StatusWord 0x60B9:
     Bit 0  Touch Probe 1 enabled
     Bit 1  Rising-edge data captured
     Bit 2  Falling-edge data captured

   IMPROVEMENT vs Confa: added tCaptureTimeout so states 20/30
   don't wait forever if the trigger never fires.
   ============================================================ *)

FUNCTION_BLOCK SML_TouchProbe
VAR_IN_OUT
    Axis : OpenSML_Axis;
END_VAR
VAR_INPUT
    xEnable          : BOOL;
    xExecute         : BOOL;          // Level: enable Touch Probe hardware
    xRisingCapture   : BOOL;          // Level: arm rising-edge latch; hold to keep result
    xFallingCapture  : BOOL;          // Level: arm falling-edge latch; hold to keep result
    xReset           : BOOL;
    tEnableTimeout   : TIME := T#200MS; // Max wait for TouchProbe_StatusWord.0 to confirm
    tCaptureTimeout  : TIME := T#5S;    // Max wait for trigger edge to arrive (0=no timeout)
END_VAR
VAR_OUTPUT
    xDone_R                  : BOOL;
    xDone_F                  : BOOL;
    xBusy                    : BOOL;
    xError                   : BOOL;
    TouchProbe_Rising_Value  : DINT; // Latched position at rising edge [encoder counts]
    TouchProbe_Falling_Value : DINT; // Latched position at falling edge [encoder counts]
    eProgress                : E_PROGRESS; // Level A: unified progress (projection of iState)
END_VAR
VAR
    iState     : INT;
    tonEnable  : TON; // Waits for probe hardware to confirm enabled
    tonCapture : TON; // Guards against trigger never arriving
END_VAR

// -- Enable/disable Touch Probe hardware every cycle -----------------------
IF xExecute AND NOT xError THEN
    Axis.TouchProbe_ControlWord.0 := TRUE;  // Enable
    Axis.TouchProbe_ControlWord.1 := FALSE; // Single-shot
    Axis.TouchProbe_ControlWord.2 := FALSE; // Trigger: DI13
ELSE
    Axis.TouchProbe_ControlWord.0 := FALSE;
    Axis.TouchProbe_ControlWord.1 := FALSE;
    Axis.TouchProbe_ControlWord.2 := FALSE;
END_IF

CASE iState OF

    0: // Idle - wait for drive ready and probe hardware enabled
        xDone_R := FALSE; xDone_F := FALSE;
        xBusy   := FALSE; xError  := FALSE;
        TouchProbe_Rising_Value  := 0;
        TouchProbe_Falling_Value := 0;

        // Timer: guard in case drive never confirms TouchProbe enabled
        tonEnable(
            IN := xExecute AND Axis.StatusWord.1 AND Axis.StatusWord.2
                  AND NOT Axis.StatusWord.3 AND Axis.StatusWord.4
                  AND NOT Axis.TouchProbe_StatusWord.0,
            PT := tEnableTimeout);

        IF xEnable THEN
            IF xExecute AND Axis.StatusWord.1 AND Axis.StatusWord.2
               AND NOT Axis.StatusWord.3 AND Axis.StatusWord.4
               AND Axis.TouchProbe_StatusWord.0 THEN
                // Drive confirmed Touch Probe 1 enabled
                tonEnable.IN := FALSE;
                iState := 10;
            ELSIF (xExecute AND tonEnable.Q) OR Axis.StatusWord.3 THEN
                iState := 999;
            END_IF
        END_IF

    10: // Armed - wait for rising or falling capture request
        IF Axis.StatusWord.3 OR NOT xEnable THEN
            iState := 999;
        ELSIF xRisingCapture THEN
            Axis.TouchProbe_ControlWord.4 := TRUE; // Arm rising-edge latch
            xBusy := TRUE;
            tonCapture.IN := FALSE;
            iState := 20;
        ELSIF xFallingCapture THEN
            Axis.TouchProbe_ControlWord.5 := TRUE; // Arm falling-edge latch
            xBusy := TRUE;
            tonCapture.IN := FALSE;
            iState := 30;
        ELSIF NOT xExecute OR NOT Axis.TouchProbe_StatusWord.0 THEN
            Axis.TouchProbe_ControlWord.4 := FALSE;
            Axis.TouchProbe_ControlWord.5 := FALSE;
            iState := 0;
        END_IF

    20: // Wait for rising-edge trigger
        // Capture timeout: if trigger never arrives, error (skip if tCaptureTimeout=0)
        tonCapture(IN := TRUE,
                   PT := SEL(tCaptureTimeout = T#0S, tCaptureTimeout, T#999999S));

